--- program FrameL_C (robot ABB IRB 1300-10/1.15) ---
  Smooth(1)
  Set speed (1000.0 mm/s)
  Set Ref.: FrameL
  Set Tool: Generic Paint Sprayer
  Show Generic Paint Sprayer
  MoveJ 1 to (-1015.17, 960.31, 527.51) mm, rotated rx -115.53 ry -8.78 rz 162.28 deg; joints [74.023, 64.389, -177.634, 4.007, 86.75, 96.944, 1374.27, 3638.377, 370.799]
  MoveL 2 to (-1015.17, 960.31, 527.51) mm, rotated rx -115.53 ry -8.78 rz 162.28 deg; joints [74.023, 64.389, -177.634, 4.007, 86.75, 96.944, 1374.27, 3638.377, 370.799]
  MoveL 3 to (-1048.89, 876.36, 484.92) mm, rotated rx -115.53 ry -8.78 rz 162.28 deg; joints [74.023, 64.389, -177.634, 4.007, 86.75, 96.944, 1340.546, 3554.421, 413.392]
  MoveL 4 to (-1048.89, 876.36, 484.92) mm, rotated rx -115.53 ry -8.78 rz 162.28 deg; joints [74.023, 64.389, -177.634, 4.007, 86.75, 96.944, 1340.546, 3554.421, 413.392]
  Set speed (200.0 mm/s)
  MoveL 5 to (-1060.66, 876.62, 493.81) mm, rotated rx -115.95 ry -8.86 rz 162.43 deg; joints [74.023, 64.389, -177.634, 3.86, 86.355, 97.028, 1327.85, 3552.819, 401.035]
  MoveL 6 to (-1082.9, 876.62, 508.72) mm, rotated rx -117.21 ry -8.2 rz 164.5 deg; joints [74.023, 64.389, -177.634, 1.62, 85.639, 97.385, 1285.601, 3546.469, 378.721]
  MoveL 7 to (-1106.18, 876.62, 522.33) mm, rotated rx -120.93 ry -8.21 rz 166.59 deg; joints [74.023, 64.389, -177.634, -0.649, 82.446, 98.449, 1245.481, 3527.612, 337.393]
  MoveL 8 to (-1130.25, 876.36, 534.1) mm, rotated rx -123.9 ry -7.79 rz 168.6 deg; joints [74.023, 64.389, -177.635, -2.986, 80.093, 99.537, 1203.573, 3510.479, 305.654]
  MoveL 9 to (-1155.11, 876.1, 544.57) mm, rotated rx -126.6 ry -7.43 rz 170.12 deg; joints [74.023, 64.389, -179.794, -4.819, 80.083, 100.454, 1169.34, 3480.642, 285.56]
  MoveL 10 to (-1181.01, 875.83, 553.72) mm, rotated rx -129.64 ry -6.78 rz 171.9 deg; joints [74.023, 64.389, -182.144, -7.096, 80.08, 101.523, 1130.972, 3446.46, 267.382]
  MoveL 11 to (-1207.43, 875.31, 561.05) mm, rotated rx -132.01 ry -6.08 rz 173.29 deg; joints [74.023, 64.389, -183.913, -8.986, 80.08, 102.381, 1093.829, 3419.143, 254.394]
  MoveL 12 to (-1234.64, 874.79, 567.06) mm, rotated rx -134.1 ry -4.52 rz 175.35 deg; joints [74.023, 64.389, -185.084, -11.889, 80.08, 103.395, 1045.347, 3394.777, 245.717]
  MoveL 13 to (-1262.63, 874, 571.51) mm, rotated rx -135.78 ry -3.02 rz 177.06 deg; joints [74.023, 64.389, -185.959, -14.438, 80.08, 104.298, 998.548, 3373.942, 240.221]
  MoveL 14 to (-1290.62, 873.22, 574.39) mm, rotated rx -136.93 ry -1.36 rz 178.73 deg; joints [74.023, 64.389, -186.309, -16.976, 80.08, 105.132, 950.472, 3358.614, 238.296]
  MoveL 15 to (-1319.14, 872.43, 575.44) mm, rotated rx -138.23 ry 0.47 rz -179.58 deg; joints [74.023, 64.389, -186.628, -19.701, 79.974, 106.138, 900.949, 3341.306, 238.296]
  MoveL 16 to (-1347.65, 871.65, 574.39) mm, rotated rx -138.48 ry 3.29 rz -177.09 deg; joints [74.023, 64.389, -185.749, -23.502, 79.974, 107.295, 839.31, 3332.647, 245.735]
  MoveL 17 to (-1375.91, 870.6, 571.77) mm, rotated rx -138.43 ry 4.69 rz -175.85 deg; joints [74.023, 64.389, -185.157, -25.368, 79.974, 107.882, 794.724, 3328.918, 252.198]
  MoveL 18 to (-1403.9, 869.82, 567.06) mm, rotated rx -137.68 ry 7.29 rz -173.41 deg; joints [74.023, 64.389, -183.479, -28.797, 79.974, 108.923, 735.673, 3328.843, 265.904]
  MoveL 19 to (-1431.63, 868.77, 560.79) mm, rotated rx -136.77 ry 8.45 rz -172.14 deg; joints [74.023, 64.389, -182.957, -30.295, 80.608, 108.944, 693.869, 3328.843, 280.789]
  MoveL 20 to (-1458.84, 867.46, 552.68) mm, rotated rx -135.42 ry 10.6 rz -169.72 deg; joints [74.023, 64.389, -181.504, -33.244, 81.1, 109.501, 640.229, 3328.841, 301.523]
  MoveL 21 to (-1485.52, 866.15, 542.73) mm, rotated rx -133.88 ry 12.26 rz -167.55 deg; joints [74.023, 64.389, -180.635, -35.596, 82.031, 109.501, 592.858, 3327.208, 325.646]
  MoveL 22 to (-1511.42, 864.59, 530.96) mm, rotated rx -131.7 ry 14.03 rz -164.78 deg; joints [74.023, 64.389, -179.236, -38.372, 82.988, 109.462, 542.722, 3327.208, 354.62]
  MoveL 23 to (-1536.8, 862.75, 517.62) mm, rotated rx -129.53 ry 15.12 rz -162.45 deg; joints [74.023, 64.389, -178.191, -40.401, 83.978, 109.007, 499.686, 3327.208, 383.586]
  MoveL 24 to (-1560.87, 860.92, 502.71) mm, rotated rx -126.89 ry 16.3 rz -159.49 deg; joints [74.023, 64.389, -176.645, -42.942, 84.889, 108.635, 454.489, 3327.209, 416.346]
  MoveL 25 to (-1585.98, 858.31, 484.39) mm, rotated rx -125.12 ry 16.78 rz -157.68 deg; joints [74.023, 64.389, -175.535, -44.366, 85.349, 108.344, 417.425, 3327.209, 445.194]
  Set speed (1000.0 mm/s)
  MoveL 26 to (-1585.98, 858.31, 484.39) mm, rotated rx -125.12 ry 16.78 rz -157.68 deg; joints [74.023, 64.389, -175.535, -44.366, 85.349, 108.344, 417.425, 3327.209, 445.194]
  MoveL 27 to (-1632.41, 927.67, 539.47) mm, rotated rx -125.12 ry 16.78 rz -157.68 deg; joints [74.023, 64.389, -175.535, -44.366, 85.349, 108.344, 371.003, 3396.571, 390.114]
  Set speed (1000.0 mm/s)
  MoveL 28 to (-1782.13, 744.91, 885.74) mm, rotated rx -119.9 ry 6.95 rz -168.12 deg; joints [74.023, 82.832, -189.902, -29.809, 83.081, 103.224, 291.65, 3396.571, 197.643]
  MoveL 29 to (-1758.39, 661.31, 836.26) mm, rotated rx -119.9 ry 6.95 rz -168.12 deg; joints [74.023, 82.832, -189.902, -29.809, 83.081, 103.224, 315.396, 3312.976, 247.119]
  MoveL 30 to (-1758.39, 661.31, 836.26) mm, rotated rx -119.9 ry 6.95 rz -168.12 deg; joints [74.023, 82.832, -189.902, -29.809, 83.081, 103.224, 315.396, 3312.976, 247.119]
  Set speed (200.0 mm/s)
  MoveL 31 to (-1724.9, 670.47, 838.1) mm, rotated rx -121.18 ry 6.48 rz -169.44 deg; joints [74.023, 82.832, -191.204, -28.584, 83.081, 103.236, 361.581, 3315.861, 237.578]
  MoveL 32 to (-1691.68, 677.53, 839.67) mm, rotated rx -120.38 ry 5.33 rz -171 deg; joints [74.023, 82.942, -191.204, -26.541, 83.271, 102.399, 409.246, 3336.803, 237.579]
  MoveL 33 to (-1652.17, 686.16, 839.67) mm, rotated rx -120.13 ry 5.09 rz -171.3 deg; joints [74.023, 82.942, -191.058, -26.131, 83.271, 102.232, 451.408, 3349.272, 237.987]
  MoveL 34 to (-1610.05, 694.54, 839.67) mm, rotated rx -119.87 ry 4.65 rz -171.96 deg; joints [74.023, 82.942, -191.057, -25.301, 83.343, 101.933, 499.698, 3362.547, 237.986]
  MoveL 35 to (-1562.18, 702.65, 839.67) mm, rotated rx -119.38 ry 4.09 rz -172.77 deg; joints [74.023, 82.942, -190.802, -24.26, 83.343, 101.565, 554.808, 3378.986, 238.548]
  MoveL 36 to (-1528.43, 707.88, 839.4) mm, rotated rx -119.36 ry 3.58 rz -173.66 deg; joints [74.023, 82.942, -190.956, -23.231, 83.343, 101.335, 597.012, 3388.041, 237.249]
  MoveL 37 to (-1485.26, 713.63, 838.88) mm, rotated rx -118.87 ry 2.94 rz -174.68 deg; joints [74.023, 82.942, -190.736, -21.967, 83.343, 100.942, 649.473, 3402.601, 238.129]
  MoveL 38 to (-1441.83, 719.13, 838.1) mm, rotated rx -117.68 ry 2.67 rz -174.93 deg; joints [74.023, 82.942, -189.774, -21.484, 83.343, 100.534, 693.898, 3420.583, 243.983]
  MoveL 39 to (-1401.81, 723.58, 837.57) mm, rotated rx -117.2 ry 2.44 rz -175.26 deg; joints [74.023, 82.942, -189.426, -21.034, 83.343, 100.319, 736.495, 3430.885, 246.249]
  MoveL 40 to (-1370.15, 726.98, 837.05) mm, rotated rx -116.96 ry 2.24 rz -175.61 deg; joints [74.023, 82.942, -189.285, -20.596, 83.343, 100.172, 771.246, 3437.889, 247.356]
  MoveL 41 to (-1348.7, 729.07, 836.53) mm, rotated rx -116.25 ry 1.82 rz -176.31 deg; joints [74.023, 82.942, -188.793, -19.705, 83.343, 99.816, 798.461, 3449.363, 250.333]
  MoveL 42 to (-1313.64, 732.47, 835.74) mm, rotated rx -115.78 ry 1.8 rz -176.28 deg; joints [74.023, 82.942, -188.382, -19.671, 83.343, 99.686, 832.592, 3457.166, 253.563]
  MoveL 43 to (-1272.05, 736.66, 834.7) mm, rotated rx -115.78 ry 1.8 rz -176.28 deg; joints [74.023, 82.942, -188.382, -19.671, 83.343, 99.686, 874.188, 3461.352, 254.61]
  Set speed (1000.0 mm/s)
  MoveL 44 to (-1272.05, 736.66, 834.7) mm, rotated rx -115.78 ry 1.8 rz -176.28 deg; joints [74.023, 82.942, -188.382, -19.671, 83.343, 99.686, 874.188, 3461.352, 254.61]
  MoveL 45 to (-1279.25, 826.43, 878.16) mm, rotated rx -115.78 ry 1.8 rz -176.28 deg; joints [74.023, 82.942, -188.382, -19.671, 83.343, 99.686, 866.984, 3551.122, 211.142]
  Set speed (1000.0 mm/s)
  MoveL 46 to (-1224.09, 625.8, 1224.25) mm, rotated rx -153.49 ry 17.59 rz -171.43 deg; joints [74.023, 113.295, -210, -50.489, 58.121, 141.888, 800.056, 3107.358, 0]
  MoveL 47 to (-1190.69, 585.7, 1138.95) mm, rotated rx -153.49 ry 17.59 rz -171.43 deg; joints [74.023, 113.295, -210, -50.489, 58.121, 141.888, 833.458, 3067.258, 85.301]
  MoveL 48 to (-1190.69, 585.7, 1138.95) mm, rotated rx -153.49 ry 17.59 rz -171.43 deg; joints [74.023, 113.295, -210, -50.489, 58.121, 141.888, 833.458, 3067.258, 85.301]
  Set speed (200.0 mm/s)
  MoveL 49 to (-1213.18, 590.41, 1127.7) mm, rotated rx -152.92 ry 17.68 rz -171.17 deg; joints [74.109, 113.295, -209.797, -50.489, 58.34, 141.571, 810.153, 3076.307, 98.867]
  MoveL 50 to (-1232.02, 595.91, 1115.67) mm, rotated rx -149.63 ry 20.03 rz -168.65 deg; joints [74.109, 113.295, -209.797, -51.349, 61.878, 139.926, 770.209, 3087.414, 138.308]
  MoveL 51 to (-1245.36, 601.66, 1104.16) mm, rotated rx -144.68 ry 22.57 rz -164.79 deg; joints [74.109, 113.295, -209.797, -52.484, 66.425, 137.222, 731.825, 3098.93, 187.325]
  MoveL 52 to (-1255.57, 608.2, 1091.34) mm, rotated rx -138.48 ry 23.76 rz -160.37 deg; joints [74.109, 113.295, -209.797, -53.093, 70.737, 133.096, 702.117, 3113.993, 238.067]
  MoveL 53 to (-1266.03, 615.79, 1076.43) mm, rotated rx -135.62 ry 23.47 rz -158.71 deg; joints [74.355, 113.295, -209.797, -53.093, 72.19, 130.762, 689.721, 3129.009, 266.528]
  MoveL 54 to (-1277.02, 624.69, 1059.16) mm, rotated rx -132.74 ry 23.27 rz -156.85 deg; joints [74.355, 113.295, -209.797, -53.171, 73.8, 128.56, 673.065, 3142.176, 298.917]
  MoveL 55 to (-1289.58, 634.63, 1039.02) mm, rotated rx -131.52 ry 23.24 rz -155.98 deg; joints [74.355, 113.295, -209.797, -53.335, 74.526, 127.689, 657.589, 3152.866, 325.984]
  MoveL 56 to (-1302.66, 645.09, 1016.52) mm, rotated rx -130.52 ry 22.58 rz -155.81 deg; joints [74.946, 113.295, -209.797, -53.335, 74.692, 126.502, 651.96, 3170.749, 350.648]
  MoveL 57 to (-1314.95, 656.34, 992.97) mm, rotated rx -127.95 ry 21.97 rz -154.38 deg; joints [75.07, 113.295, -209.797, -53.335, 75.943, 124.315, 637.676, 3187.198, 386.491]
  MoveL 58 to (-1325.16, 667.33, 969.69) mm, rotated rx -124.78 ry 21.2 rz -152.49 deg; joints [75.07, 113.295, -209.797, -53.423, 77.573, 121.661, 622.718, 3202.179, 425.966]
  MoveL 59 to (-1331.7, 677.01, 948.5) mm, rotated rx -121.28 ry 19.57 rz -151.13 deg; joints [75.729, 113.295, -209.797, -53.423, 78.977, 118.19, 621.847, 3223.413, 462.069]
  MoveL 60 to (-1334.83, 686.16, 929.14) mm, rotated rx -115.7 ry 16.94 rz -148.81 deg; joints [76.214, 113.295, -209.797, -53.423, 81.501, 112.732, 620.29, 3244.805, 508.191]
  MoveL 61 to (-1335.36, 694.54, 911.09) mm, rotated rx -112.21 ry 15.04 rz -147.57 deg; joints [76.419, 113.295, -209.796, -53.344, 83.103, 109.182, 620.29, 3260.09, 543.538]
  MoveL 62 to (-1334.05, 702.65, 894.34) mm, rotated rx -108.35 ry 12.58 rz -146.71 deg; joints [76.419, 113.295, -208.835, -52.795, 84.285, 105.811, 620.291, 3284.293, 577.893]
  MoveL 63 to (-1330.91, 710.23, 878.65) mm, rotated rx -106.25 ry 11.06 rz -146.65 deg; joints [76.419, 113.295, -207.305, -52.247, 84.285, 104.649, 622.688, 3310.154, 601.765]
  MoveL 64 to (-1326.72, 717.82, 863.73) mm, rotated rx -104 ry 9.39 rz -146.81 deg; joints [76.419, 113.295, -205.674, -51.514, 84.285, 103.354, 626.889, 3338.129, 626.047]
  MoveL 65 to (-1321.23, 725.14, 849.35) mm, rotated rx -102.7 ry 8.13 rz -147.88 deg; joints [76.419, 113.295, -204.934, -50.104, 84.286, 102.209, 637.653, 3363.4, 645.188]
  MoveL 66 to (-1354.46, 721.74, 850.39) mm, rotated rx -175.54 ry 33.28 rz 101.98 deg; joints [56.988, 143.589, -137.16, 144.417, 41.145, 36.117, 651.946, 3698.807, 1100]
  MoveL 67 to (-1365.71, 720.44, 850.65) mm, rotated rx -146.28 ry 2.17 rz -178.55 deg; joints [76.42, 113.126, -204.934, -34.5, 46.983, 127.515, 802.993, 3345.808, 316.76]
  MoveL 68 to (-1402.07, 716.25, 851.7) mm, rotated rx -146.28 ry 2.15 rz -178.57 deg; joints [76.452, 113.127, -204.934, -34.5, 46.968, 127.491, 767.195, 3341.791, 315.632]
  MoveL 69 to (-1441.57, 711.54, 852.75) mm, rotated rx -147.29 ry 2.97 rz -178.09 deg; joints [76.452, 113.127, -205.051, -36.188, 46.968, 129.159, 719.979, 3326.698, 313.434]
  MoveL 70 to (-1483.95, 705.52, 854.05) mm, rotated rx -147.72 ry 2.66 rz -178.32 deg; joints [76.657, 113.126, -205.225, -36.188, 46.589, 129.171, 683.277, 3317.897, 308.963]
  MoveL 71 to (-1526.07, 699.25, 855.1) mm, rotated rx -148.75 ry 3.4 rz -177.94 deg; joints [76.657, 113.126, -205.394, -37.74, 46.589, 130.742, 634.518, 3301.013, 306.662]
  MoveL 72 to (-1565.32, 692.97, 855.89) mm, rotated rx -149.59 ry 4.5 rz -177.37 deg; joints [76.657, 113.076, -205.394, -39.637, 46.907, 132.518, 585.134, 3285.408, 306.662]
  MoveL 73 to (-1604.04, 685.64, 856.67) mm, rotated rx -149.63 ry 4.75 rz -177.22 deg; joints [76.657, 113.053, -205.394, -39.955, 47.091, 132.754, 544.052, 3276.943, 306.662]
  MoveL 74 to (-1644.85, 677.27, 857.19) mm, rotated rx -149.67 ry 5.03 rz -177.07 deg; joints [76.657, 112.983, -205.394, -40.272, 47.328, 132.968, 500.693, 3267.189, 306.662]
  MoveL 75 to (-1683.3, 668.64, 857.72) mm, rotated rx -149.88 ry 4.86 rz -177.19 deg; joints [76.768, 112.983, -205.475, -40.272, 47.126, 132.968, 465.246, 3257.352, 304.541]
  MoveL 76 to (-1714.44, 661.05, 857.72) mm, rotated rx -150.07 ry 5.32 rz -176.94 deg; joints [76.768, 112.823, -205.475, -40.855, 47.48, 133.411, 429.986, 3246.468, 304.541]
  MoveL 77 to (-1699.79, 652.15, 878.91) mm, rotated rx -108.33 ry -41.93 rz 178.16 deg; joints [107.262, 119.949, -159.707, -81.239, 23.985, 121.042, 1096.293, 3778.444, 604.845]
  MoveL 78 to (-1684.35, 642.74, 900.88) mm, rotated rx -103.77 ry -3.13 rz 167.42 deg; joints [76.148, 112.823, -205.475, -3.654, 79.163, 94.041, 621.106, 3510.146, 535.977]
  MoveL 79 to (-1667.87, 633.06, 924.17) mm, rotated rx -103.52 ry -3.2 rz 166.93 deg; joints [76.148, 113.008, -205.475, -3.137, 79.163, 93.889, 642.032, 3502.509, 516.04]
  MoveL 80 to (-1650.34, 622.85, 949.02) mm, rotated rx -103.61 ry -3.24 rz 166.87 deg; joints [76.148, 113.007, -205.475, -3.08, 79.072, 93.904, 660.131, 3492.212, 490.338]
  MoveL 81 to (-1668.13, 617.1, 950.85) mm, rotated rx -150.18 ry 3.36 rz -178.08 deg; joints [76.148, 127.331, -159.488, -126.409, 33.343, 234.838, 410.502, 3521.9, 490.338]
  MoveL 82 to (-1646.94, 607.16, 976.49) mm, rotated rx -103.2 ry -21.92 rz 173.54 deg; joints [79.337, 132.004, -146.722, -134.913, 10.128, 208.962, 623.21, 3814.134, 838.601]
  MoveL 83 to (-1626.27, 597.74, 1000.82) mm, rotated rx -103.03 ry 17 rz 164.34 deg; joints [83.994, 114.805, -210, -10.723, 92.781, 110.214, 765.634, 3467.741, 546.847]
  MoveL 84 to (-1604.3, 587.54, 1026.46) mm, rotated rx -102.27 ry -2.64 rz 168.02 deg; joints [68.793, 127.331, -142.872, 39.964, 4.671, 54.643, 479.375, 3792.466, 820.793]
  MoveL 85 to (-1591.22, 581.26, 1041.37) mm, rotated rx -102.7 ry -2.7 rz 168.18 deg; joints [68.793, 127.33, -143.048, 40.106, 4.387, 54.643, 491.326, 3784.586, 800.784]
  MoveL 86 to (-1576.3, 574.19, 1058.38) mm, rotated rx -102.74 ry -2.72 rz 168.15 deg; joints [68.821, 127.318, -143.074, 40.113, 4.387, 54.643, 506.991, 3777.652, 783.064]
  MoveL 87 to (-1558.25, 565.82, 1078.78) mm, rotated rx -102.36 ry -3.02 rz 166.5 deg; joints [69.84, 127.318, -143.735, 40.113, 5.465, 54.375, 557.879, 3777.653, 760.069]
  MoveL 88 to (-1552.24, 562.68, 1085.58) mm, rotated rx -103.74 ry -3.73 rz 165.11 deg; joints [71.265, 127.318, -145.275, 40.29, 5.465, 54.375, 602.999, 3777.836, 728.411]
  MoveL 89 to (-1529.74, 549.6, 1110.17) mm, rotated rx -104.95 ry -3.95 rz 165.55 deg; joints [71.265, 127.318, -145.818, 40.635, 4.699, 54.375, 622.506, 3759.732, 689.247]
  MoveL 90 to (-1522.15, 545.15, 1118.55) mm, rotated rx -106.77 ry -4.5 rz 165.41 deg; joints [71.357, 127.318, -147.645, 41.199, 4.699, 54.375, 636.151, 3745.82, 651.363]
  MoveL 91 to (-1514.83, 540.71, 1126.66) mm, rotated rx -108.15 ry -4.97 rz 165.21 deg; joints [71.531, 127.318, -149.051, 41.589, 4.699, 54.375, 650.887, 3734.192, 620.842]
  MoveL 92 to (-1509.07, 536.52, 1132.93) mm, rotated rx -109.08 ry -4.93 rz 166.05 deg; joints [71.623, 127.66, -149.051, 41.589, 3.22, 54.557, 650.887, 3725.698, 612.176]
  MoveL 93 to (-1479.25, 539.4, 1137.12) mm, rotated rx -96.71 ry 0.66 rz -174.4 deg; joints [52.115, 127.659, -135.62, 39.626, 3.22, 54.557, 184.512, 3559.834, 826.74]
  MoveL 94 to (-1446.02, 542.02, 1141.57) mm, rotated rx -96.9 ry 0.66 rz -174.6 deg; joints [52.293, 127.659, -135.786, 39.725, 3.22, 54.557, 222.003, 3564.9, 819.431]
  MoveL 95 to (-1405.47, 545.15, 1147.32) mm, rotated rx -96.24 ry 0.57 rz -174.82 deg; joints [52.145, 127.685, -135.786, 39.725, 3.877, 54.18, 262.446, 3568.064, 819.43]
  MoveL 96 to (-1359.69, 548.56, 1153.34) mm, rotated rx -95.72 ry 0.46 rz -175.39 deg; joints [52.145, 127.685, -136.116, 39.725, 4.814, 53.897, 313.297, 3574.124, 815.026]
  MoveL 97 to (-1311.03, 551.96, 1159.88) mm, rotated rx -93.84 ry 0.28 rz -175.81 deg; joints [51.521, 127.643, -136.116, 38.704, 6.754, 53.892, 356.743, 3574.124, 823.22]
  MoveL 98 to (-1261.84, 555.1, 1165.9) mm, rotated rx -94.32 ry 0.29 rz -176.15 deg; joints [51.809, 127.643, -136.507, 38.986, 6.754, 53.892, 413.141, 3581.111, 810.29]
  MoveL 99 to (-1215.02, 557.97, 1171.39) mm, rotated rx -92.6 ry 0.13 rz -177.14 deg; joints [51.285, 127.075, -136.507, 38.986, 9.273, 53.02, 459.516, 3585.376, 810.29]
  MoveL 100 to (-1166.36, 560.59, 1176.62) mm, rotated rx -90.9 ry 0.05 rz -177.14 deg; joints [50.926, 127.075, -135.847, 37.989, 10.12, 53.02, 502.442, 3585.376, 824.087]
  MoveL 101 to (-1111.42, 562.94, 1181.86) mm, rotated rx -88.74 ry -0.04 rz -178.11 deg; joints [50.117, 126.225, -135.847, 37.074, 13.323, 52.861, 552.192, 3585.376, 824.096]
  MoveL 102 to (-1049.68, 565.56, 1187.09) mm, rotated rx -86.59 ry -0.11 rz -178.18 deg; joints [49.822, 126.225, -134.979, 35.766, 14.298, 52.861, 609.4, 3585.372, 843.363]
  MoveL 103 to (-981.39, 567.91, 1192.32) mm, rotated rx -85.14 ry -0.19 rz -177.72 deg; joints [49.495, 126.224, -133.896, 34.792, 14.298, 52.861, 668.023, 3582.496, 858.047]
  MoveL 104 to (-904.48, 570.79, 1197.55) mm, rotated rx -82.67 ry -0.17 rz -178.69 deg; joints [48.935, 125.631, -133.896, 33.479, 17.36, 52.86, 743.872, 3582.496, 864.961]
  MoveL 105 to (-818.15, 573.41, 1202.52) mm, rotated rx -79.46 ry -0.27 rz -178.56 deg; joints [48.899, 125.631, -131.755, 31.359, 17.672, 52.86, 826.261, 3582.495, 902.412]
  MoveL 106 to (-727.89, 576.29, 1206.71) mm, rotated rx -76.16 ry -0.16 rz -179.35 deg; joints [48.815, 125.631, -130.971, 29.412, 19.77, 52.86, 921.427, 3582.494, 932.118]
  MoveL 107 to (-639.73, 578.9, 1209.85) mm, rotated rx -75.2 ry -0.12 rz -179.54 deg; joints [48.665, 125.631, -130.915, 28.851, 20.562, 52.86, 1009.092, 3582.084, 937.49]
  MoveL 108 to (-560.72, 581.26, 1212.2) mm, rotated rx -74.25 ry -0.19 rz -179.34 deg; joints [48.251, 125.631, -130.748, 28.203, 21.141, 52.86, 1080.603, 3576.71, 943.985]
  MoveL 109 to (-498.72, 583.09, 1213.25) mm, rotated rx -72.59 ry -0.34 rz -178.92 deg; joints [47.368, 125.631, -130.664, 27.035, 22.339, 52.86, 1126.833, 3562.073, 956.627]
  MoveL 110 to (-447.18, 584.66, 1213.25) mm, rotated rx -73.06 ry -0.49 rz -178.38 deg; joints [47.122, 125.631, -130.664, 27.035, 21.798, 53.038, 1170.327, 3559.537, 952.194]
  MoveL 111 to (-400.61, 585.97, 1212.73) mm, rotated rx -72.12 ry -0.65 rz -177.98 deg; joints [46.48, 125.631, -130.66, 26.321, 22.465, 53.038, 1204.822, 3548.789, 959.813]
  MoveL 112 to (-356.92, 587.54, 1211.94) mm, rotated rx -70.24 ry -0.72 rz -177.99 deg; joints [45.923, 125.631, -130.659, 25.065, 23.969, 53.038, 1241.071, 3538.165, 975.631]
  MoveL 113 to (-315.06, 588.84, 1210.63) mm, rotated rx -70.43 ry -0.9 rz -177.46 deg; joints [45.525, 125.631, -130.659, 25.049, 23.68, 53.038, 1273.107, 3532.715, 974.676]
  MoveL 114 to (-272.42, 590.41, 1208.8) mm, rotated rx -70.97 ry -0.97 rz -177.19 deg; joints [45.384, 125.631, -130.79, 25.348, 23.331, 53.038, 1311.73, 3532.716, 970.896]
  MoveL 115 to (-226.9, 591.98, 1206.45) mm, rotated rx -73.64 ry -0.96 rz -176.74 deg; joints [44.998, 125.631, -132.354, 27.122, 22.863, 53.038, 1350.313, 3532.716, 940.01]
  MoveL 116 to (-177.19, 594.08, 1203.57) mm, rotated rx -73.35 ry -0.99 rz -176.7 deg; joints [44.899, 125.631, -132.32, 26.914, 23.048, 53.038, 1398.384, 3532.716, 945.435]
  MoveL 117 to (-122.25, 596.95, 1199.65) mm, rotated rx -71 ry -1.16 rz -176.62 deg; joints [44.814, 125.631, -130.978, 25.227, 23.367, 53.038, 1449.764, 3529.34, 977.622]
  MoveL 118 to (-64.7, 600.35, 1194.68) mm, rotated rx -71.58 ry -1.55 rz -175.36 deg; joints [43.91, 125.631, -130.978, 25.227, 22.594, 53.107, 1484.953, 3516.791, 976.338]
  MoveL 119 to (-7.41, 604.28, 1188.4) mm, rotated rx -71.84 ry -2 rz -173.91 deg; joints [42.65, 125.483, -130.978, 25.042, 22.207, 53.107, 1513.724, 3498.226, 976.338]
  MoveL 120 to (47.53, 608.73, 1180.55) mm, rotated rx -71.95 ry -2.25 rz -173.12 deg; joints [41.878, 125.238, -130.978, 24.927, 22.207, 53.107, 1551.811, 3489.375, 978.496]
  MoveL 121 to (97.76, 613.17, 1171.39) mm, rotated rx -72.14 ry -2.58 rz -172.05 deg; joints [40.827, 124.881, -130.978, 24.806, 22.207, 53.107, 1579.348, 3475.469, 979.235]
  MoveL 122 to (146.16, 618.14, 1160.67) mm, rotated rx -71.66 ry -3.12 rz -170.66 deg; joints [39.492, 124.881, -130.973, 24.071, 22.208, 53.107, 1600.414, 3453.1, 991.733]
  MoveL 123 to (195.08, 623.9, 1148.11) mm, rotated rx -70.72 ry -3.9 rz -168.99 deg; joints [37.886, 124.881, -130.779, 22.861, 22.208, 53.107, 1616.753, 3424.083, 1010.129]
  MoveL 124 to (244.27, 630.96, 1132.67) mm, rotated rx -72.37 ry -4.39 rz -166.45 deg; joints [36.316, 124.881, -130.779, 22.861, 20.403, 53.762, 1629.557, 3398.061, 1010.086]
  MoveL 125 to (293.45, 639.6, 1113.05) mm, rotated rx -73.81 ry -4.79 rz -163.94 deg; joints [34.487, 124.485, -130.779, 22.861, 19.275, 54.345, 1640.022, 3368.784, 1010.086]
  MoveL 126 to (347.34, 650.58, 1088.98) mm, rotated rx -75.56 ry -4.41 rz -163.38 deg; joints [33.9, 124.103, -131.5, 24.28, 19.275, 54.345, 1684.493, 3372.016, 1010.086]
  MoveL 127 to (411.18, 663.4, 1059.94) mm, rotated rx -77.83 ry -3.62 rz -163.67 deg; joints [34.059, 123.592, -132.235, 26.347, 19.275, 54.345, 1752.616, 3394.507, 1010.086]
  MoveL 128 to (478.41, 677.27, 1028.03) mm, rotated rx -76.13 ry -4.13 rz -163.75 deg; joints [33.354, 123.589, -132.235, 25.979, 20.539, 53.289, 1812.432, 3394.507, 1054.104]
  MoveL 129 to (541.98, 690.61, 996.11) mm, rotated rx -77.3 ry -3.78 rz -163.69 deg; joints [32.777, 122.082, -132.235, 27.086, 21.487, 53.29, 1865.951, 3404.149, 1054.105]
  MoveL 130 to (598.49, 702.38, 966.55) mm, rotated rx -81.33 ry -2.4 rz -164.67 deg; joints [33.246, 122.082, -134.352, 30.848, 21.487, 53.29, 1939.65, 3433.922, 1040.16]
  MoveL 131 to (643.49, 711.8, 942.22) mm, rotated rx -81.55 ry -2.4 rz -164.23 deg; joints [32.765, 121.878, -134.352, 30.997, 21.523, 53.29, 1976.214, 3433.922, 1059.38]
  MoveL 132 to (682.21, 719.91, 920.5) mm, rotated rx -82.28 ry -2.2 rz -164.16 deg; joints [32.181, 120.834, -134.352, 31.735, 22.267, 53.29, 2006.381, 3435.187, 1059.38]
  MoveL 133 to (719.36, 727.76, 899.05) mm, rotated rx -81.72 ry -2.4 rz -163.96 deg; joints [31.793, 120.699, -134.352, 31.309, 22.767, 53.248, 2037.804, 3435.187, 1082.681]
  MoveL 134 to (754.41, 735.09, 878.65) mm, rotated rx -79.11 ry -3.34 rz -163.15 deg; joints [31.295, 117.378, -129.937, 28.826, 23.013, 53.248, 2045.276, 3435.187, 1100]
  MoveL 135 to (786.59, 741.63, 859.03) mm, rotated rx -81.68 ry -2.48 rz -163.48 deg; joints [31.207, 117.378, -131.27, 31.246, 23.013, 53.248, 2082.657, 3444.94, 1091.877]
  MoveL 136 to (817.2, 748.17, 839.93) mm, rotated rx -80.71 ry -2.91 rz -162.77 deg; joints [30.689, 115.081, -128.534, 30.247, 23.013, 53.248, 2093.261, 3443.042, 1100]
  MoveL 137 to (846.24, 754.18, 821.61) mm, rotated rx -82.59 ry -2.12 rz -164.12 deg; joints [31.66, 115.081, -129.394, 32.148, 23.013, 53.248, 2143.77, 3474.649, 1099.433]
  MoveL 138 to (874.76, 760.2, 803.3) mm, rotated rx -81.97 ry -2.36 rz -163.7 deg; joints [31.181, 112.683, -126.999, 31.58, 23.359, 53.248, 2156.086, 3474.648, 1100]
  Set speed (1000.0 mm/s)
  MoveL 139 to (874.76, 760.2, 803.3) mm, rotated rx -81.97 ry -2.36 rz -163.7 deg; joints [31.181, 112.683, -126.999, 31.58, 23.359, 53.248, 2156.086, 3474.648, 1100]
  MoveL 140 to (846.41, 855.08, 789.34) mm, rotated rx -81.97 ry -2.36 rz -163.7 deg; joints [30.702, 111.825, -126.999, 31.58, 24.332, 53.381, 2122.171, 3562.297, 1100]
  Set speed (1000.0 mm/s)
  MoveL 141 to (1541.36, 940.82, 613.61) mm, rotated rx -125.26 ry -7.23 rz 169.91 deg; joints [30.702, 111.825, -161.462, 74.993, 31.83, 53.381, 3191.702, 3594.263, 705.738]
  MoveL 142 to (1519.9, 861.71, 556.34) mm, rotated rx -125.26 ry -7.23 rz 169.91 deg; joints [30.702, 111.825, -161.462, 74.992, 31.83, 53.381, 3170.245, 3515.153, 763.012]
  MoveL 143 to (1519.9, 861.71, 556.34) mm, rotated rx -125.26 ry -7.23 rz 169.91 deg; joints [30.702, 111.825, -161.462, 74.992, 31.83, 53.381, 3170.245, 3515.153, 763.012]
  Set speed (200.0 mm/s)
  MoveL 144 to (1494, 861.45, 566.8) mm, rotated rx -125.78 ry -6.92 rz 170.51 deg; joints [30.702, 112.149, -161.462, 74.964, 31.003, 53.381, 3137.514, 3511.708, 754.412]
  MoveL 145 to (1489.29, 872.43, 551.89) mm, rotated rx -123.78 ry -6.41 rz 170.52 deg; joints [29.063, 112.149, -160.887, 74.915, 33.272, 53.381, 3113.809, 3511.71, 787.542]
  MoveL 146 to (1461.56, 872.96, 561.57) mm, rotated rx -124.95 ry -6.3 rz 171.08 deg; joints [29.508, 112.243, -160.887, 75.006, 31.785, 53.381, 3084.564, 3511.71, 771.24]
  MoveL 147 to (1433.04, 873.48, 569.68) mm, rotated rx -126.07 ry -5.47 rz 172.55 deg; joints [29.508, 113.123, -160.887, 74.89, 29.817, 53.381, 3039.121, 3504.629, 770.22]
  MoveL 148 to (1404.52, 874.26, 576.22) mm, rotated rx -127.67 ry -4.4 rz 174.32 deg; joints [29.608, 114.1, -160.812, 74.89, 27.168, 53.381, 2990.793, 3495.601, 770.22]
  MoveL 149 to (1375.22, 875.05, 580.67) mm, rotated rx -128.32 ry -3.5 rz 175.58 deg; joints [29.609, 114.229, -159.976, 74.684, 25.574, 53.381, 2943.185, 3492.131, 770.22]
  MoveL 150 to (1345.92, 876.1, 583.81) mm, rotated rx -128.52 ry -2.35 rz 177.05 deg; joints [29.609, 114.229, -158.608, 74.132, 24.01, 53.381, 2890.52, 3491.681, 776.48]
  MoveL 151 to (1316.1, 876.88, 585.12) mm, rotated rx -127.31 ry -1.42 rz 178.14 deg; joints [29.1, 114.229, -157.227, 73.229, 24.008, 53.381, 2837.13, 3491.681, 793.636]
  MoveL 152 to (1286.01, 877.67, 585.38) mm, rotated rx -125.42 ry -0.49 rz 179.31 deg; joints [28.402, 114.229, -155.682, 71.968, 24.501, 53.381, 2781.001, 3491.681, 817.801]
  MoveL 153 to (1255.14, 878.45, 584.07) mm, rotated rx -122.83 ry 0.38 rz -179.41 deg; joints [27.568, 114.229, -154.001, 70.247, 25.437, 53.381, 2722.233, 3491.682, 849.706]
  MoveL 154 to (1223.49, 879.24, 581.45) mm, rotated rx -120.01 ry 0.77 rz -178.66 deg; joints [26.72, 114.229, -152.909, 68.545, 27.094, 53.381, 2671.668, 3491.684, 880.366]
  MoveL 155 to (1190.26, 879.5, 578.05) mm, rotated rx -117.18 ry 1.29 rz -177.49 deg; joints [26.075, 114.229, -151.527, 66.485, 28.178, 53.381, 2616.373, 3491.684, 914.661]
  MoveL 156 to (1155.47, 879.5, 573.87) mm, rotated rx -116.01 ry 1.07 rz -177.82 deg; joints [26.075, 114.16, -151.527, 65.79, 29.242, 53.381, 2584.953, 3497.655, 925.992]
  MoveL 157 to (1117.01, 879.24, 569.16) mm, rotated rx -111.18 ry 0.83 rz -177.85 deg; joints [24.971, 114.161, -151.225, 63.037, 33.256, 53.381, 2537.979, 3497.655, 969.43]
  MoveL 158 to (1107.07, 868.25, 594.8) mm, rotated rx -116 ry 0.51 rz -178.95 deg; joints [26.602, 114.161, -152.303, 65.955, 29.946, 53.381, 2554.828, 3497.655, 898.648]
  MoveL 159 to (1106.28, 861.97, 607.09) mm, rotated rx -118.35 ry 0.15 rz -179.73 deg; joints [27.54, 114.16, -153.145, 67.339, 28.498, 53.381, 2572.558, 3497.655, 862.408]
  MoveL 160 to (1067.3, 855.17, 619.65) mm, rotated rx -120.95 ry -0.25 rz 179.58 deg; joints [28.69, 114.16, -154.04, 68.676, 26.683, 53.381, 2553.898, 3497.655, 824.139]
  MoveL 161 to (1017.6, 845.23, 638.48) mm, rotated rx -122.6 ry -1.12 rz 178.25 deg; joints [29.774, 114.16, -155.4, 69.641, 26.174, 53.381, 2533.298, 3497.655, 782.834]
  MoveL 162 to (977.57, 845.23, 640.58) mm, rotated rx -121.89 ry -1.11 rz 178.22 deg; joints [29.525, 114.16, -155.285, 69.349, 26.819, 53.381, 2490.792, 3497.658, 786.521]
  MoveL 163 to (935.97, 845.23, 643.19) mm, rotated rx -121.07 ry -1.09 rz 178.19 deg; joints [29.243, 114.16, -155.155, 69, 27.567, 53.381, 2446.403, 3497.658, 790.674]
  MoveL 164 to (924.99, 833.19, 664.12) mm, rotated rx -120.71 ry -1.09 rz 178.17 deg; joints [29.523, 114.331, -155.154, 68.587, 27.563, 53.381, 2437.619, 3491.47, 774.824]
  MoveL 165 to (917.4, 825.08, 678.25) mm, rotated rx -120.01 ry -1.07 rz 178.15 deg; joints [29.835, 114.949, -155.154, 68.534, 27.625, 52.692, 2432.154, 3491.47, 774.824]
  MoveL 166 to (912.43, 820.11, 687.93) mm, rotated rx -118.12 ry -1.03 rz 178.08 deg; joints [29.552, 114.949, -154.763, 67.478, 29.028, 52.692, 2423.355, 3491.494, 781.508]
  MoveL 167 to (907.98, 815.92, 696.56) mm, rotated rx -117.18 ry -1 rz 178.05 deg; joints [29.536, 114.97, -154.56, 66.865, 29.626, 52.692, 2417.985, 3491.495, 781.508]
  MoveL 168 to (945.13, 815.66, 693.69) mm, rotated rx -117.42 ry -1.01 rz 178.05 deg; joints [29.536, 114.896, -154.56, 66.994, 29.486, 52.723, 2455.16, 3490.236, 781.508]
  MoveL 169 to (982.02, 815.4, 690.81) mm, rotated rx -117.89 ry -1.02 rz 178.07 deg; joints [29.696, 114.896, -154.623, 67.203, 29.06, 52.723, 2493.6, 3490.236, 780.424]
  MoveL 170 to (1018.91, 815.14, 688.19) mm, rotated rx -118.36 ry -1.23 rz 177.73 deg; joints [29.832, 114.896, -155.009, 67.591, 29.016, 52.723, 2536.911, 3490.235, 776.618]
  MoveL 171 to (1056.05, 814.62, 685.31) mm, rotated rx -119.54 ry -1.67 rz 177.06 deg; joints [30.199, 114.896, -155.82, 68.447, 28.69, 52.723, 2587.894, 3490.23, 764.715]
  MoveL 172 to (1094.51, 814.09, 682.17) mm, rotated rx -120.25 ry -1.69 rz 177.1 deg; joints [30.472, 114.896, -155.921, 68.72, 28.018, 52.723, 2628.94, 3490.229, 761.976]
  MoveL 173 to (1134.8, 813.31, 678.77) mm, rotated rx -120.96 ry -1.71 rz 177.15 deg; joints [30.769, 114.896, -156.022, 68.974, 27.328, 52.723, 2672.03, 3490.229, 759.546]
  MoveL 174 to (1177.97, 812.52, 674.85) mm, rotated rx -121.67 ry -2.16 rz 176.51 deg; joints [31.045, 114.896, -156.75, 69.55, 27.334, 52.723, 2727.821, 3490.229, 752.808]
  MoveL 175 to (1222.44, 811.48, 670.66) mm, rotated rx -121.68 ry -2.37 rz 176.17 deg; joints [31.073, 114.693, -156.846, 69.689, 27.649, 52.723, 2776.774, 3490.229, 752.808]
  MoveL 176 to (1266.65, 810.43, 666.22) mm, rotated rx -121.92 ry -2.59 rz 175.86 deg; joints [31.218, 114.666, -157.142, 69.894, 27.703, 52.723, 2827.021, 3490.229, 752.808]
  MoveL 177 to (1308.77, 809.12, 661.51) mm, rotated rx -124.52 ry -2.92 rz 175.77 deg; joints [32.313, 114.666, -157.886, 70.872, 25.463, 52.723, 2884.542, 3490.151, 733.89]
  MoveL 178 to (1347.49, 807.81, 657.32) mm, rotated rx -125.02 ry -3.6 rz 174.87 deg; joints [32.613, 114.666, -158.852, 71.389, 25.852, 52.723, 2940.606, 3490.151, 727.32]
  MoveL 179 to (1385.95, 806.24, 652.35) mm, rotated rx -125.03 ry -3.83 rz 174.56 deg; joints [32.686, 114.384, -158.852, 71.49, 26.104, 52.723, 2983.535, 3490.151, 727.478]
  MoveL 180 to (1427.28, 804.15, 646.59) mm, rotated rx -125.23 ry -4.17 rz 174.12 deg; joints [32.909, 114.274, -159.19, 71.666, 26.266, 52.723, 3033.678, 3490.151, 727.478]
  MoveL 181 to (1486.67, 800.49, 637.18) mm, rotated rx -126.06 ry -5.23 rz 172.86 deg; joints [33.603, 114.274, -160.59, 72.301, 26.528, 52.723, 3120.904, 3490.151, 720.778]
  MoveL 182 to (1530.1, 797.35, 629.59) mm, rotated rx -125.49 ry -5.54 rz 172.29 deg; joints [33.55, 113.974, -160.59, 72.269, 27.436, 52.723, 3170.153, 3490.151, 727.159]
  MoveL 183 to (1571.43, 793.43, 622) mm, rotated rx -126.36 ry -6.17 rz 171.7 deg; joints [33.678, 113.974, -161.534, 73.024, 27.436, 52.723, 3225.026, 3481.37, 722.239]
  MoveL 184 to (1603.09, 790.02, 615.99) mm, rotated rx -125.07 ry -7.05 rz 170.09 deg; joints [33.678, 113.109, -161.582, 73.087, 29.648, 52.723, 3275.022, 3486.215, 722.239]
  MoveL 185 to (1632.65, 786.1, 609.97) mm, rotated rx -121.53 ry -6.97 rz 168.82 deg; joints [32.468, 113.109, -161.33, 72.481, 33.588, 52.723, 3301.948, 3486.215, 754.871]
  MoveL 186 to (1604.14, 786.62, 621.48) mm, rotated rx -118.75 ry -5.87 rz 169.45 deg; joints [31.246, 113.109, -159.904, 71.212, 35.486, 52.723, 3245.588, 3486.216, 774.116]
  Set speed (1000.0 mm/s)
  MoveL 187 to (1604.14, 786.62, 621.48) mm, rotated rx -118.75 ry -5.87 rz 169.45 deg; joints [31.246, 113.109, -159.904, 71.212, 35.486, 52.723, 3245.588, 3486.216, 774.116]
  MoveL 188 to (1625.03, 871.91, 669.33) mm, rotated rx -118.75 ry -5.87 rz 169.45 deg; joints [31.246, 113.109, -159.904, 71.212, 35.486, 52.723, 3266.48, 3571.502, 726.265]
  Set speed (1000.0 mm/s)
  MoveL 189 to (944.76, 961.41, 628.52) mm, rotated rx -102.53 ry -0.15 rz 179.33 deg; joints [22.48, 113.109, -152.046, 60.314, 43.621, 52.723, 2378.942, 3571.502, 957.472]
  MoveL 190 to (943.56, 863.8, 606.83) mm, rotated rx -102.53 ry -0.15 rz 179.33 deg; joints [22.48, 113.109, -152.046, 60.314, 43.621, 52.723, 2377.738, 3473.892, 979.167]
  MoveL 191 to (943.56, 863.8, 606.83) mm, rotated rx -102.53 ry -0.15 rz 179.33 deg; joints [22.48, 113.109, -152.046, 60.314, 43.621, 52.723, 2377.738, 3473.892, 979.167]
  Set speed (200.0 mm/s)
  MoveL 192 to (941.47, 865.37, 600.81) mm, rotated rx -103.3 ry -0.03 rz 179.89 deg; joints [22.48, 113.109, -152.046, 60.227, 42.743, 53.164, 2370.668, 3471.796, 979.259]
  MoveL 193 to (942.51, 867.72, 592.44) mm, rotated rx -104.82 ry 0.09 rz -179.67 deg; joints [22.635, 113.379, -152.046, 60.966, 41.175, 53.192, 2368.53, 3471.796, 979.256]
  MoveL 194 to (948.53, 871.13, 580.67) mm, rotated rx -104.47 ry 0.2 rz -179.23 deg; joints [22.461, 113.379, -151.846, 60.518, 41.165, 53.274, 2368.53, 3471.796, 995.471]
  MoveL 195 to (961.35, 877.14, 557.65) mm, rotated rx -101.65 ry 0.35 rz -178.31 deg; joints [21.918, 113.379, -151.344, 58.304, 42.654, 53.274, 2367.518, 3471.796, 1045.45]
  MoveL 196 to (968.94, 884.47, 522.07) mm, rotated rx -98.82 ry 0.38 rz -177.58 deg; joints [21.394, 113.036, -151.344, 55.674, 44.685, 53.957, 2366.085, 3471.796, 1100]
  MoveL 197 to (959.52, 887.08, 495.38) mm, rotated rx -96 ry 0.33 rz -176.86 deg; joints [21.363, 109.565, -151.344, 50.43, 48.362, 58.052, 2355.854, 3471.797, 1100]
  MoveL 198 to (949.84, 888.13, 477.07) mm, rotated rx -93.88 ry 0.21 rz -176.84 deg; joints [21.342, 107.078, -151.344, 47.67, 51.524, 60.107, 2351.553, 3471.796, 1100]
  MoveL 199 to (939.64, 888.39, 457.97) mm, rotated rx -92.71 ry 0.15 rz -176.83 deg; joints [21.429, 105.064, -151.344, 45.847, 53.719, 61.731, 2347.453, 3471.796, 1100]
  MoveL 200 to (929.69, 888.65, 437.83) mm, rotated rx -92 ry 0.11 rz -176.83 deg; joints [21.49, 103.237, -151.344, 44.523, 55.502, 63.165, 2343.762, 3470.933, 1100]
  MoveL 201 to (920.8, 888.65, 416.9) mm, rotated rx -90.71 ry 0.04 rz -176.82 deg; joints [21.49, 100.987, -151.344, 42.933, 58.101, 64.627, 2343.161, 3467.92, 1099.993]
  MoveL 202 to (912.69, 888.13, 394.4) mm, rotated rx -89.41 ry -0.04 rz -176.35 deg; joints [21.49, 98.6, -151.344, 40.968, 60.666, 66.288, 2341.199, 3461.341, 1100]
  MoveL 203 to (905.89, 887.61, 373.21) mm, rotated rx -88.94 ry -0.08 rz -175.41 deg; joints [21.49, 96.782, -151.344, 39.168, 62.052, 67.912, 2335.131, 3453.109, 1100]
  MoveL 204 to (900.66, 886.82, 356.2) mm, rotated rx -88.24 ry -0.14 rz -175.42 deg; joints [21.49, 94.919, -150.64, 38.552, 63.497, 68.439, 2335.131, 3450.131, 1100]
  MoveL 205 to (895.95, 886.04, 340.77) mm, rotated rx -88.24 ry -0.14 rz -175.42 deg; joints [21.49, 93.7, -150.334, 38.273, 64.212, 69.071, 2335.131, 3447.494, 1100]
  Set speed (1000.0 mm/s)
  MoveL 206 to (895.95, 886.04, 340.77) mm, rotated rx -88.24 ry -0.14 rz -175.42 deg; joints [21.49, 93.7, -150.334, 38.273, 64.212, 69.071, 2335.131, 3447.494, 1100]
  MoveL 207 to (887.95, 985.67, 337.69) mm, rotated rx -88.24 ry -0.14 rz -175.42 deg; joints [21.425, 93.472, -150.334, 38.273, 64.413, 69.196, 2328.017, 3545.651, 1100]
  Set speed (1000.0 mm/s)
  MoveL 208 to (853.38, 969.89, 348.17) mm, rotated rx -103.01 ry 7.43 rz -150.75 deg; joints [21.425, 93.472, -150.334, 9.922, 49.835, 97.581, 2115.612, 3359.096, 994.29]
  MoveL 209 to (903.53, 886.3, 325.86) mm, rotated rx -103.01 ry 7.43 rz -150.75 deg; joints [21.425, 93.472, -150.334, 9.922, 49.835, 97.581, 2165.763, 3275.508, 1016.606]
  MoveL 210 to (903.53, 886.3, 325.86) mm, rotated rx -103.01 ry 7.43 rz -150.75 deg; joints [21.425, 93.472, -150.334, 9.922, 49.835, 97.581, 2165.763, 3275.508, 1016.606]
  Set speed (200.0 mm/s)
  MoveL 211 to (914.52, 887.87, 345.22) mm, rotated rx -100.5 ry 6.57 rz -148.31 deg; joints [22.118, 93.472, -149.767, 6.474, 50.738, 97.381, 2165.763, 3275.326, 1016.606]
  MoveL 212 to (923.42, 888.65, 365.1) mm, rotated rx -102.16 ry 7.09 rz -150.22 deg; joints [21.962, 93.472, -149.766, 8.81, 49.725, 97.381, 2182.992, 3285.205, 984.925]
  MoveL 213 to (934.14, 889.44, 387.07) mm, rotated rx -103.41 ry 7.4 rz -151.62 deg; joints [21.92, 93.472, -149.767, 10.449, 48.952, 97.381, 2200.549, 3293.301, 953.912]
  MoveL 214 to (946.44, 890.22, 410.1) mm, rotated rx -105.74 ry 8.32 rz -152.83 deg; joints [21.683, 93.472, -149.758, 11.746, 47.568, 98.672, 2216.557, 3293.302, 915.548]
  MoveL 215 to (959.78, 890.48, 431.55) mm, rotated rx -108.87 ry 9.31 rz -154.67 deg; joints [21.399, 93.472, -149.758, 13.694, 45.669, 100.099, 2236.545, 3293.302, 872.978]
  MoveL 216 to (974.43, 890.75, 451.95) mm, rotated rx -110.73 ry 9.77 rz -155.85 deg; joints [21.224, 93.472, -149.758, 14.989, 44.51, 100.768, 2255.807, 3293.302, 839.728]
  MoveL 217 to (990.13, 890.48, 471.05) mm, rotated rx -114.55 ry 10.34 rz -158.54 deg; joints [20.905, 93.472, -149.758, 18.008, 42.046, 101.659, 2283.287, 3293.302, 793.397]
  MoveL 218 to (1011.58, 890.22, 492.77) mm, rotated rx -108.25 ry 10.08 rz -152.05 deg; joints [20.905, 93.472, -149.758, 10.729, 46.351, 102.075, 2270.138, 3267.055, 820.098]
  MoveL 219 to (1023.61, 888.13, 515.53) mm, rotated rx -113.08 ry 11.73 rz -154.49 deg; joints [20.905, 94.219, -149.758, 12.318, 42.718, 105.094, 2287.457, 3267.055, 776.725]
  Set speed (1000.0 mm/s)
  MoveL 220 to (1023.61, 888.13, 515.53) mm, rotated rx -113.08 ry 11.73 rz -154.49 deg; joints [20.905, 94.219, -149.758, 12.318, 42.718, 105.094, 2287.457, 3267.055, 776.725]
  MoveL 221 to (976.81, 967.73, 553.91) mm, rotated rx -113.08 ry 11.73 rz -154.49 deg; joints [20.905, 94.219, -149.758, 12.318, 42.718, 105.094, 2240.65, 3346.653, 738.343]

--- program FrameR_C (robot ABB IRB 1300-10/1.15) ---
  Smooth(1)
  Set speed (1000.0 mm/s)
  Set Ref.: FrameR
  Set Tool: Generic Paint Sprayer
  Show Generic Paint Sprayer
  MoveJ 1 to (-1567.41, -947.44, 561.3) mm, rotated rx 116.18 ry 8.07 rz 164.06 deg; joints [-18.613, 70.643, -160.975, 159.818, -72.367, 68.936, 14.365, 240.215, 405.979]
  MoveL 2 to (-1567.41, -947.44, 561.3) mm, rotated rx 116.18 ry 8.07 rz 164.06 deg; joints [-18.613, 70.643, -160.975, 159.818, -72.367, 68.936, 14.365, 240.215, 405.979]
  MoveL 3 to (-1536.8, -862.85, 517.62) mm, rotated rx 116.18 ry 8.07 rz 164.06 deg; joints [-18.613, 70.643, -160.975, 159.818, -72.367, 68.936, 44.975, 324.8, 449.664]
  MoveL 4 to (-1536.8, -862.85, 517.62) mm, rotated rx 116.18 ry 8.07 rz 164.06 deg; joints [-18.613, 70.643, -160.975, 159.818, -72.367, 68.936, 44.975, 324.8, 449.664]
  Set speed (200.0 mm/s)
  MoveL 5 to (-1511.42, -864.68, 530.96) mm, rotated rx 117.6 ry 7.57 rz 165.86 deg; joints [-18.613, 70.643, -160.975, 158.345, -70.921, 68.501, 83.279, 316.894, 423.259]
  MoveL 6 to (-1485.52, -866.25, 542.73) mm, rotated rx 119.49 ry 6.77 rz 168.23 deg; joints [-18.613, 70.643, -160.989, 156.392, -68.942, 68.006, 127.136, 308.433, 393.799]
  MoveL 7 to (-1458.84, -867.56, 552.68) mm, rotated rx 120.63 ry 6.22 rz 169.63 deg; joints [-18.608, 70.645, -160.989, 155.208, -67.701, 67.76, 164.896, 303.689, 373.04]
  MoveL 8 to (-1431.63, -868.61, 560.79) mm, rotated rx 121.87 ry 5.07 rz 171.91 deg; joints [-18.608, 70.645, -161.394, 153.058, -66.382, 67.76, 214.467, 295.937, 351.142]
  MoveL 9 to (-1403.9, -869.65, 567.06) mm, rotated rx 122.48 ry 4.46 rz 173.04 deg; joints [-18.608, 70.645, -161.65, 151.982, -65.747, 67.76, 254.1, 292.049, 337.984]
  MoveL 10 to (-1375.91, -870.7, 571.77) mm, rotated rx 122.85 ry 3.63 rz 174.4 deg; joints [-18.607, 70.645, -162.511, 150.654, -65.699, 67.76, 300.795, 287.554, 327.831]
  MoveL 11 to (-1347.65, -871.48, 574.39) mm, rotated rx 123.43 ry 2.18 rz 176.71 deg; joints [-18.607, 70.645, -163.965, 148.372, -65.568, 67.76, 361.589, 281.477, 316.442]
  MoveL 12 to (-1319.14, -872.53, 575.44) mm, rotated rx 123.01 ry 1.1 rz 178.31 deg; joints [-18.607, 70.645, -164.386, 146.346, -65.568, 68.646, 409.222, 272.173, 314.488]
  MoveL 13 to (-1290.62, -873.32, 574.39) mm, rotated rx 122.75 ry 0.03 rz 179.95 deg; joints [-18.607, 70.645, -164.966, 144.398, -65.568, 69.295, 458.433, 264.711, 313.88]
  MoveL 14 to (-1262.63, -874.1, 571.51) mm, rotated rx 121.5 ry -0.87 rz -178.58 deg; joints [-18.607, 70.645, -164.966, 142.218, -65.996, 70.794, 501.334, 252.628, 322.32]
  MoveL 15 to (-1234.64, -874.62, 567.06) mm, rotated rx 119.59 ry -1.16 rz -177.95 deg; joints [-18.607, 70.645, -164.966, 140.919, -67.366, 72.2, 535.411, 241.481, 339.756]
  MoveL 16 to (-1207.43, -875.41, 561.05) mm, rotated rx 117.47 ry -1.89 rz -176.36 deg; joints [-18.607, 70.645, -164.966, 138.54, -68.641, 74.029, 577.946, 226.627, 358.999]
  MoveL 17 to (-1181.01, -875.67, 553.72) mm, rotated rx 114.97 ry -2.36 rz -174.95 deg; joints [-18.607, 70.645, -164.966, 136.4, -70.403, 75.823, 617.522, 212.418, 383.818]
  MoveL 18 to (-1155.11, -876.19, 544.57) mm, rotated rx 113.17 ry -2.69 rz -173.75 deg; joints [-18.607, 70.645, -164.966, 134.745, -71.68, 77.07, 654.392, 202.078, 405.856]
  MoveL 19 to (-1130.25, -876.46, 534.1) mm, rotated rx 110.41 ry -2.6 rz -173.06 deg; joints [-18.607, 70.645, -164.966, 133.557, -74.022, 78.489, 684.783, 190.934, 438.633]
  MoveL 20 to (-1106.18, -876.46, 522.33) mm, rotated rx 107.69 ry -2.35 rz -172.66 deg; joints [-18.607, 70.645, -164.966, 132.771, -76.442, 79.73, 711.467, 182.061, 473.425]
  MoveL 21 to (-1082.9, -876.72, 508.72) mm, rotated rx 105 ry -2.28 rz -171.55 deg; joints [-18.607, 70.645, -164.966, 131.287, -78.713, 81.041, 744.285, 172.206, 509.473]
  MoveL 22 to (-1060.66, -876.46, 493.81) mm, rotated rx 102.34 ry -1.62 rz -172.64 deg; joints [-18.368, 70.645, -164.966, 131.892, -81.381, 81.898, 754.662, 172.209, 549.165]
  MoveL 23 to (-1048.89, -876.46, 484.92) mm, rotated rx 101.61 ry -1.74 rz -171.59 deg; joints [-18.368, 70.645, -164.966, 130.744, -81.892, 82.332, 775.999, 168.058, 563.788]
  Set speed (1000.0 mm/s)
  MoveL 24 to (-1048.89, -876.46, 484.92) mm, rotated rx 101.61 ry -1.74 rz -171.59 deg; joints [-18.368, 70.645, -164.966, 130.744, -81.892, 82.332, 775.999, 168.058, 563.788]
  MoveL 25 to (-1033.96, -973.27, 505.03) mm, rotated rx 101.61 ry -1.74 rz -171.59 deg; joints [-18.368, 70.645, -164.966, 130.744, -81.892, 82.332, 790.935, 71.246, 543.68]
  Set speed (1000.0 mm/s)
  MoveL 26 to (-1620.34, -905.96, 635.31) mm, rotated rx 95.09 ry -1.66 rz -161.98 deg; joints [-23.506, 70.645, -168.71, 125.797, -89.471, 82.332, 337.544, 71.246, 474.728]
  MoveL 27 to (-1651.39, -811.31, 626.45) mm, rotated rx 95.09 ry -1.66 rz -161.98 deg; joints [-23.507, 70.645, -168.71, 125.798, -89.471, 82.332, 306.493, 165.888, 483.588]
  MoveL 28 to (-1651.39, -811.31, 626.45) mm, rotated rx 95.09 ry -1.66 rz -161.98 deg; joints [-23.507, 70.645, -168.71, 125.798, -89.471, 82.332, 306.493, 165.888, 483.588]
  Set speed (200.0 mm/s)
  MoveL 29 to (-1645.89, -808.17, 640.32) mm, rotated rx 113.53 ry -8.08 rz -162.12 deg; joints [-23.507, 72.673, -168.71, 127.007, -69.184, 79.927, 306.494, 206.634, 309.416]
  MoveL 30 to (-1651.65, -799.02, 663.34) mm, rotated rx 121.42 ry -9.52 rz -164.85 deg; joints [-23.507, 72.673, -168.71, 130.57, -61.954, 76.902, 284.437, 252.951, 222.205]
  MoveL 31 to (-1666.56, -784.63, 693.42) mm, rotated rx 124.61 ry -9.92 rz -165.99 deg; joints [-23.507, 73.957, -168.71, 131.64, -58.294, 76.527, 250.715, 279.424, 178.795]
  MoveL 32 to (-1677.55, -774.95, 712.52) mm, rotated rx 126.3 ry -10.62 rz -165.92 deg; joints [-23.574, 73.957, -168.71, 131.661, -56.497, 76.164, 244.342, 297.996, 145.936]
  MoveL 33 to (-1683.83, -769.72, 722.72) mm, rotated rx 125.13 ry -10.25 rz -165.82 deg; joints [-23.558, 73.957, -169.107, 131.661, -57.93, 76.164, 239.386, 297.902, 145.355]
  MoveL 34 to (-1683.83, -769.72, 722.72) mm, rotated rx 171.16 ry 2.79 rz 179.57 deg; joints [-36.296, 73.957, -189.291, 194.827, -57.93, 27.33, 239.385, 619.77, 42.153]
  MoveL 35 to (-1643.8, -776.52, 722.72) mm, rotated rx 171.27 ry 13.42 rz 177.96 deg; joints [-36.914, 73.957, -189.291, 200.842, -67.394, 24.825, 197.215, 619.774, 96.315]
  MoveL 36 to (-1607.96, -779.4, 730.31) mm, rotated rx 167.94 ry 10.28 rz 177.82 deg; joints [-33.158, 73.957, -189.291, 194.194, -66.22, 26.961, 238.044, 614.627, 76.195]
  MoveL 37 to (-1574.47, -782.8, 735.54) mm, rotated rx 162.76 ry 12.18 rz 176.26 deg; joints [-33.158, 73.957, -186.255, 192.105, -66.997, 30.46, 238.043, 566.815, 81.388]
  Set speed (1000.0 mm/s)
  MoveL 38 to (-1574.47, -782.8, 735.54) mm, rotated rx 162.76 ry 12.18 rz 176.26 deg; joints [-33.158, 73.957, -186.255, 192.105, -66.997, 30.46, 238.043, 566.815, 81.388]
  MoveL 39 to (-1596.51, -811.05, 828.9) mm, rotated rx 162.76 ry 12.18 rz 176.26 deg; joints [-33.158, 75.195, -187.492, 192.105, -66.997, 30.46, 213.238, 536.755, 0.003]
  Set speed (1000.0 mm/s)
  MoveL 40 to (-1593.63, -878.91, 757.51) mm, rotated rx 98.12 ry 1.45 rz 169.97 deg; joints [-33.158, 75.195, -183.445, 163.358, -101.211, 79.486, 213.238, 138.256, 406.615]
  MoveL 41 to (-1576.04, -781.49, 743.39) mm, rotated rx 98.12 ry 1.45 rz 169.97 deg; joints [-33.158, 75.195, -183.445, 163.358, -101.211, 79.486, 230.829, 235.678, 420.735]
  MoveL 42 to (-1576.04, -781.49, 743.39) mm, rotated rx 98.12 ry 1.45 rz 169.97 deg; joints [-33.158, 75.195, -183.445, 163.358, -101.211, 79.486, 230.829, 235.678, 420.735]
  Set speed (200.0 mm/s)
  MoveL 43 to (-1574.47, -782.27, 739.73) mm, rotated rx 97.18 ry 1.28 rz 169.93 deg; joints [-33.158, 75.195, -183.201, 163.264, -101.701, 80.152, 230.829, 233.1, 431.046]
  MoveL 44 to (-1571.6, -783.32, 735.54) mm, rotated rx 102.36 ry 2.06 rz 170.68 deg; joints [-33.158, 75.729, -183.201, 163.488, -97.124, 76.98, 234.295, 233.103, 398.064]
  MoveL 45 to (-1568.19, -785.41, 730.05) mm, rotated rx 108.49 ry 2.67 rz 172.07 deg; joints [-33.158, 76.713, -183.201, 163.595, -91.261, 73.401, 239.31, 233.102, 362.103]
  MoveL 46 to (-1563.75, -789.08, 722.2) mm, rotated rx 111.32 ry 2.84 rz 172.75 deg; joints [-33.158, 76.962, -183.201, 163.705, -88.725, 71.728, 246.486, 233.102, 349.55]
  MoveL 47 to (-1557.21, -794.31, 711.74) mm, rotated rx 113.21 ry 2.87 rz 173.35 deg; joints [-33.158, 76.962, -183.201, 163.673, -87.145, 70.589, 257.356, 231.07, 345.118]
  MoveL 48 to (-1543.86, -806.08, 689.5) mm, rotated rx 112.74 ry 3 rz 172.89 deg; joints [-32.822, 76.962, -182.72, 163.673, -87.145, 70.89, 262.386, 220.973, 370.252]
  MoveL 49 to (-1538.37, -810.27, 681.65) mm, rotated rx 112.52 ry 3.31 rz 172.07 deg; joints [-32.75, 76.961, -182.72, 164.391, -87.566, 70.949, 260.5, 220.973, 381.211]
  MoveL 50 to (-1531.83, -814.19, 674.59) mm, rotated rx 113.2 ry 2.69 rz 173.74 deg; joints [-32.75, 76.961, -182.72, 162.867, -86.528, 70.657, 281.259, 210.637, 380.287]
  MoveL 51 to (-1524.51, -817.85, 668.31) mm, rotated rx 113.92 ry 2.93 rz 173.42 deg; joints [-32.75, 76.961, -182.72, 163.435, -86.107, 70.178, 285.413, 211.149, 381.936]
  MoveL 52 to (-1516.4, -821.25, 663.08) mm, rotated rx 112.76 ry 3.01 rz 172.86 deg; joints [-32.542, 76.961, -182.257, 163.435, -86.681, 70.937, 285.42, 206.557, 395.395]
  MoveL 53 to (-1507.76, -824.39, 658.89) mm, rotated rx 109.21 ry 2.91 rz 171.71 deg; joints [-32.402, 76.916, -182.257, 163.435, -89.666, 73.068, 285.419, 199.674, 427.279]
  MoveL 54 to (-1498.61, -826.75, 656.01) mm, rotated rx 109.9 ry 2.54 rz 173.03 deg; joints [-32.402, 76.916, -182.258, 162.277, -88.785, 72.69, 305.443, 192.437, 423.021]
  MoveL 55 to (-1489.19, -828.84, 654.18) mm, rotated rx 107.78 ry 2.44 rz 172.43 deg; joints [-32.365, 76.916, -181.423, 162.277, -89.745, 74.227, 305.447, 184.607, 439.56]
  MoveL 56 to (-1479.51, -830.41, 653.66) mm, rotated rx 108.96 ry 2.29 rz 173.36 deg; joints [-32.365, 76.916, -181.423, 161.636, -88.611, 73.537, 322.581, 181.509, 429.869]
  MoveL 57 to (-1428.23, -836.69, 652.87) mm, rotated rx 112.95 ry 1.82 rz 175.71 deg; joints [-32.365, 76.916, -181.424, 160.346, -84.86, 71.308, 393.108, 176.138, 396.691]
  MoveL 58 to (-1385.33, -840.88, 652.09) mm, rotated rx 113.89 ry 1.35 rz 176.95 deg; joints [-32.365, 76.916, -181.424, 159.328, -83.722, 70.904, 447.029, 169.407, 388.191]
  MoveL 59 to (-1341.9, -844.02, 651.57) mm, rotated rx 113.18 ry 1.15 rz 177.32 deg; joints [-32.365, 76.916, -181.269, 158.734, -84.013, 71.415, 492.999, 161.611, 393.106]
  MoveL 60 to (-1314.69, -845.58, 651.04) mm, rotated rx 113.65 ry 1.17 rz 177.34 deg; joints [-32.249, 77.105, -181.269, 158.734, -83.449, 71.189, 518.198, 161.611, 391.36]
  MoveL 61 to (-1305.01, -845.58, 652.35) mm, rotated rx 113.89 ry 1.18 rz 177.34 deg; joints [-32.235, 77.284, -181.269, 158.773, -83.092, 71.116, 526.446, 161.611, 389.548]
  MoveL 62 to (-1296.12, -844.28, 656.27) mm, rotated rx 112.25 ry 0.44 rz 178.92 deg; joints [-32.235, 77.284, -181.226, 156.661, -83.843, 72.256, 549.803, 150.421, 395.544]
  MoveL 63 to (-1288.27, -842.18, 662.29) mm, rotated rx 109.89 ry -0.2 rz -179.46 deg; joints [-32.235, 77.284, -181.225, 154.389, -85.281, 73.661, 572.589, 138.737, 405.907]
  MoveL 64 to (-1282.25, -839.04, 669.88) mm, rotated rx 113.65 ry 0.48 rz 178.91 deg; joints [-32.235, 77.286, -181.23, 157.059, -82.712, 71.482, 563.484, 160.403, 371.001]
  MoveL 65 to (-1278.85, -835.12, 679.03) mm, rotated rx 113.65 ry 0.13 rz 179.7 deg; joints [-32.317, 77.286, -181.23, 156.309, -82.452, 71.61, 574.687, 160.404, 360.488]
  MoveL 66 to (-1277.54, -830.93, 688.71) mm, rotated rx 113.66 ry 0.65 rz 178.52 deg; joints [-32.317, 77.71, -181.23, 157.531, -82.452, 71.603, 561.67, 167.436, 355.878]
  MoveL 67 to (-1279.11, -826.49, 698.39) mm, rotated rx 113.19 ry 1.66 rz 176.12 deg; joints [-32.317, 77.959, -181.23, 159.893, -83.38, 71.634, 536.353, 179.707, 355.876]
  MoveL 68 to (-1282.51, -822.82, 706.5) mm, rotated rx 112.01 ry 1.43 rz 176.46 deg; joints [-32.317, 77.951, -181.23, 159.203, -84.202, 72.371, 536.352, 177.924, 356.114]
  MoveL 69 to (-1287.22, -818.9, 715.4) mm, rotated rx 109.18 ry 1.43 rz 175.91 deg; joints [-32.485, 77.234, -181.23, 159.196, -87.271, 73.747, 533.82, 177.924, 364.649]
  MoveL 70 to (-1291.67, -816.02, 722.99) mm, rotated rx 105.18 ry 1.04 rz 176.17 deg; joints [-32.485, 77.049, -181.23, 157.979, -90.559, 75.959, 533.82, 170.277, 387.037]
  MoveL 71 to (-1294.81, -814.45, 728.74) mm, rotated rx 100.47 ry 0.65 rz 176.47 deg; joints [-32.485, 77.049, -181.224, 156.739, -94.298, 78.535, 533.825, 161.41, 419.179]
  MoveL 72 to (-1297.16, -813.67, 732.67) mm, rotated rx 97.77 ry 0.62 rz 175.5 deg; joints [-32.485, 77.049, -181.224, 157.267, -96.675, 80.1, 523.529, 162.939, 438.079]
  MoveL 73 to (-1298.99, -813.14, 736.07) mm, rotated rx 89.91 ry -0.01 rz 175.41 deg; joints [-32.485, 76.771, -181.224, 156.398, -103.36, 84.313, 523.529, 160.679, 497.487]
  Set speed (1000.0 mm/s)
  MoveL 74 to (-1298.99, -813.14, 736.07) mm, rotated rx 89.91 ry -0.01 rz 175.41 deg; joints [-32.485, 76.771, -181.224, 156.398, -103.36, 84.313, 523.529, 160.679, 497.487]
  MoveL 75 to (-1306.99, -912.82, 735.92) mm, rotated rx 89.91 ry -0.01 rz 175.41 deg; joints [-32.485, 76.771, -181.224, 156.398, -103.36, 84.313, 515.53, 61, 497.634]
  Set speed (1000.0 mm/s)
  MoveL 76 to (-1277.26, -812.46, 899.51) mm, rotated rx 130.43 ry 1.94 rz 177.73 deg; joints [-32.485, 82.485, -181.224, 164.314, -65.405, 62.278, 515.529, 241.607, 65.66]
  MoveL 77 to (-1272.05, -736.49, 834.7) mm, rotated rx 130.43 ry 1.94 rz 177.73 deg; joints [-32.485, 82.485, -181.224, 164.314, -65.405, 62.278, 520.743, 317.58, 130.474]
  MoveL 78 to (-1272.05, -736.49, 834.7) mm, rotated rx 130.43 ry 1.94 rz 177.73 deg; joints [-32.485, 82.485, -181.224, 164.314, -65.405, 62.278, 520.743, 317.58, 130.474]
  Set speed (200.0 mm/s)
  MoveL 79 to (-1313.64, -732.57, 835.74) mm, rotated rx 131.13 ry 1.86 rz 177.87 deg; joints [-32.486, 82.485, -181.225, 164.465, -64.816, 61.836, 480.451, 324.806, 124.566]
  MoveL 80 to (-1348.7, -729.17, 836.53) mm, rotated rx 131.51 ry 2.46 rz 177.23 deg; joints [-32.486, 82.585, -181.206, 165.473, -64.817, 61.212, 437.294, 332.811, 124.566]
  MoveL 81 to (-1370.15, -726.81, 837.05) mm, rotated rx 131.03 ry 2.25 rz 177.41 deg; joints [-32.486, 82.375, -181.206, 165.02, -65.244, 61.624, 419.632, 332.534, 124.566]
  MoveL 82 to (-1401.81, -723.67, 837.57) mm, rotated rx 132.04 ry 2.5 rz 177.23 deg; joints [-32.486, 82.375, -181.206, 165.762, -64.645, 60.747, 385.483, 342.305, 118.589]
  MoveL 83 to (-1441.84, -719.23, 838.1) mm, rotated rx 133.18 ry 2.93 rz 176.89 deg; joints [-32.49, 82.375, -181.783, 166.881, -64.645, 59.499, 344.476, 357.293, 113.753]
  MoveL 84 to (-1485.26, -713.73, 838.88) mm, rotated rx 133.65 ry 3 rz 176.86 deg; joints [-32.492, 82.375, -182.089, 167.201, -64.645, 59.035, 302.34, 366.865, 110.952]
  MoveL 85 to (-1528.43, -707.71, 839.4) mm, rotated rx 134.21 ry 4.21 rz 175.68 deg; joints [-32.492, 82.375, -181.644, 169.049, -64.645, 57.959, 242.645, 380.514, 111.34]
  MoveL 86 to (-1562.18, -702.74, 839.67) mm, rotated rx 135.2 ry 4.73 rz 175.31 deg; joints [-32.493, 82.375, -181.868, 170.148, -64.51, 56.845, 205.151, 394.369, 107.799]
  MoveL 87 to (-1610.05, -694.63, 839.67) mm, rotated rx 135.22 ry 5.08 rz 174.98 deg; joints [-32.493, 82.375, -181.638, 170.602, -64.511, 56.652, 152, 403.576, 108.755]
  MoveL 88 to (-1652.17, -686.26, 839.67) mm, rotated rx 135.73 ry 5.47 rz 174.69 deg; joints [-32.493, 82.375, -181.727, 171.316, -64.511, 56.005, 106.555, 417.077, 107.647]
  MoveL 89 to (-1691.68, -677.63, 839.67) mm, rotated rx 136.03 ry 5.85 rz 174.38 deg; joints [-32.493, 82.383, -181.727, 171.926, -64.56, 55.539, 63.117, 429.319, 107.647]
  MoveL 90 to (-1724.9, -670.56, 838.1) mm, rotated rx 136.82 ry 6.43 rz 174 deg; joints [-32.493, 82.383, -181.876, 172.973, -64.56, 54.549, 25.38, 444.226, 107.518]
  MoveL 91 to (-1758.39, -661.41, 836.26) mm, rotated rx 135.23 ry 8 rz 172.14 deg; joints [-34.724, 80.46, -181.876, 176.549, -68.763, 55.099, 0.002, 444.226, 110.987]
  Set speed (1000.0 mm/s)
  MoveL 92 to (-1758.39, -661.41, 836.26) mm, rotated rx 135.23 ry 8 rz 172.14 deg; joints [-34.724, 80.46, -181.876, 176.549, -68.763, 55.099, 0.002, 444.226, 110.987]
  MoveL 93 to (-1777.81, -729.83, 906.56) mm, rotated rx 135.23 ry 8 rz 172.14 deg; joints [-34.724, 80.46, -185.22, 176.62, -72.101, 54.888, 0, 389.269, 48.578]
  Set speed (1000.0 mm/s)
  MoveL 94 to (892.89, -973.97, 160.56) mm, rotated rx 74.09 ry -79.65 rz -165.04 deg; joints [-50.625, 101.986, -183.176, 143.958, -56.047, 174.635, 2943.702, -296.83, 1100]
  MoveL 95 to (894.12, -874.1, 165.49) mm, rotated rx 74.09 ry -79.65 rz -165.04 deg; joints [-50.625, 102.249, -183.176, 143.853, -55.834, 174.822, 2944.041, -198.044, 1097.78]
  MoveL 96 to (894.12, -874.1, 165.49) mm, rotated rx 74.09 ry -79.65 rz -165.04 deg; joints [-50.625, 102.249, -183.176, 143.853, -55.834, 174.822, 2944.041, -198.044, 1097.78]
  Set speed (200.0 mm/s)
  MoveL 97 to (897.25, -874.89, 176.21) mm, rotated rx 65.87 ry -79.15 rz -157.31 deg; joints [-50.572, 102.13, -183.176, 144.306, -57.481, 174.822, 2944.041, -202.933, 1099.813]
  MoveL 98 to (899.87, -876.46, 192.17) mm, rotated rx 61.84 ry -78.73 rz -152.65 deg; joints [-50.572, 102.13, -183.176, 143.646, -58.425, 174.912, 2952.705, -207.84, 1091.736]
  MoveL 99 to (903.01, -878.29, 209.44) mm, rotated rx 62.04 ry -78.65 rz -151.92 deg; joints [-50.572, 102.13, -183.176, 142.694, -58.517, 174.948, 2963.908, -210.297, 1074.532]
  MoveL 100 to (906.93, -880.12, 229.58) mm, rotated rx 62.24 ry -78.57 rz -151.18 deg; joints [-50.572, 102.13, -183.176, 141.745, -58.61, 174.982, 2975.895, -212.626, 1054.448]
  MoveL 101 to (912.69, -881.95, 251.82) mm, rotated rx 63.48 ry -78.61 rz -151.46 deg; joints [-50.572, 102.13, -183.22, 140.789, -58.506, 174.982, 2989.943, -213.842, 1030.144]
  MoveL 102 to (920.28, -883.78, 275.36) mm, rotated rx 64.54 ry -78.72 rz -152.5 deg; joints [-50.571, 102.13, -183.221, 140.765, -58.272, 174.982, 2997.54, -214.928, 1004.496]
  MoveL 103 to (929.69, -885.35, 299.69) mm, rotated rx 65.62 ry -78.83 rz -153.56 deg; joints [-50.545, 102.13, -183.227, 140.714, -58.045, 174.982, 3006.729, -215.496, 978.065]
  MoveL 104 to (940.68, -886.66, 324.29) mm, rotated rx 66.79 ry -78.9 rz -154.23 deg; joints [-50.519, 102.13, -183.265, 140.199, -57.891, 174.982, 3021.693, -215.76, 951.388]
  MoveL 105 to (953.5, -887.97, 348.36) mm, rotated rx 85.13 ry -19.62 rz -174.48 deg; joints [0, 44.016, -168.118, 113.546, -98.533, 78.32, 3060.514, 351.718, 637.921]
  MoveL 106 to (968.15, -889.01, 371.64) mm, rotated rx 85.13 ry -19.62 rz -174.48 deg; joints [0, 44.016, -168.118, 113.546, -98.533, 78.32, 3075.164, 350.671, 614.638]
  MoveL 107 to (984.11, -889.8, 393.88) mm, rotated rx 84.63 ry -19.58 rz -174.31 deg; joints [0, 44.835, -168.118, 113.424, -98.568, 79.239, 3080.491, 349.61, 598.511]
  MoveL 108 to (1001.38, -890.32, 415.07) mm, rotated rx 85.13 ry -19.62 rz -174.48 deg; joints [0.001, 44.853, -168.118, 113.658, -98.197, 79.096, 3097.541, 349.369, 573.162]
  MoveL 109 to (1020.21, -890.58, 435.21) mm, rotated rx 84.63 ry -19.58 rz -174.31 deg; joints [0.001, 45.265, -168.118, 113.481, -98.396, 79.637, 3111.032, 348.831, 558.239]
  MoveL 110 to (1040.1, -890.84, 453.79) mm, rotated rx 84.38 ry -19.55 rz -174.23 deg; joints [0.001, 45.523, -168.118, 113.402, -98.476, 79.957, 3127.571, 348.445, 542.424]
  MoveL 111 to (1066.78, -890.84, 475.24) mm, rotated rx 84.63 ry -19.58 rz -174.31 deg; joints [0.001, 45.532, -168.118, 113.517, -98.289, 79.885, 3154.15, 348.57, 518.893]
  MoveL 112 to (1095.03, -890.58, 494.6) mm, rotated rx 85.13 ry -19.62 rz -174.48 deg; joints [0.001, 45.549, -168.118, 113.748, -97.917, 79.739, 3182.208, 349.108, 495.375]
  MoveL 113 to (1124.86, -890.06, 511.6) mm, rotated rx 85.38 ry -19.72 rz -175.5 deg; joints [0.001, 45.558, -168.118, 114.693, -98.158, 79.939, 3203.662, 352.782, 476.029]
  MoveL 114 to (1155.99, -889.54, 525.99) mm, rotated rx 85.88 ry -19.72 rz -175.19 deg; joints [0, 45.573, -168.118, 114.51, -97.577, 79.649, 3238.754, 352.115, 457.625]
  MoveL 115 to (1181.63, -888.75, 535.67) mm, rotated rx 86.12 ry -19.77 rz -175.75 deg; joints [0, 45.582, -168.118, 115.04, -97.607, 79.708, 3260.15, 354.598, 445.767]
  MoveL 116 to (1207.79, -887.97, 543.52) mm, rotated rx 86.62 ry -19.83 rz -176.38 deg; joints [0, 45.6, -168.118, 115.686, -97.454, 79.686, 3281.974, 357.321, 433.7]
  MoveL 117 to (1234.47, -887.18, 549.8) mm, rotated rx 86.87 ry -19.87 rz -176.94 deg; joints [0, 45.613, -168.118, 116.215, -97.485, 79.743, 3304.394, 359.899, 425.291]
  MoveL 118 to (1261.68, -886.4, 554.25) mm, rotated rx 87.62 ry -19.89 rz -176.72 deg; joints [0, 45.625, -168.118, 116.15, -96.728, 79.358, 3335.564, 359.768, 414.744]
  MoveL 119 to (1288.89, -885.35, 556.86) mm, rotated rx 88.12 ry -19.93 rz -177.36 deg; joints [0, 45.643, -168.118, 116.795, -96.582, 79.323, 3358.44, 362.895, 407.98]
  MoveL 120 to (1316.36, -884.57, 557.91) mm, rotated rx 88.12 ry -19.96 rz -178.3 deg; joints [0.004, 45.662, -168.118, 117.618, -97.006, 79.598, 3377.48, 366.981, 406.875]
  MoveL 121 to (1343.57, -883.78, 556.86) mm, rotated rx 88.12 ry -19.96 rz -178.3 deg; joints [0.004, 45.662, -168.118, 117.618, -97.006, 79.598, 3404.688, 367.766, 407.922]
  MoveL 122 to (1371.04, -883, 554.25) mm, rotated rx 87.87 ry -19.95 rz -178.21 deg; joints [-0.098, 45.662, -168.118, 117.592, -97.231, 79.716, 3432.156, 367.766, 412.586]
  MoveL 123 to (1398.24, -882.21, 549.8) mm, rotated rx 88.12 ry -19.96 rz -178.3 deg; joints [-0.098, 45.668, -168.118, 117.708, -97.052, 79.628, 3459.294, 368.802, 415]
  MoveL 124 to (1425.45, -881.43, 543.52) mm, rotated rx 88.87 ry -19.98 rz -178.56 deg; joints [-0.098, 45.682, -168.118, 118.055, -96.518, 79.362, 3486.317, 370.389, 415.176]
  MoveL 125 to (1452.4, -880.64, 535.67) mm, rotated rx 88.87 ry -19.98 rz -178.56 deg; joints [-0.098, 45.682, -168.118, 118.055, -96.518, 79.362, 3513.264, 371.174, 423.025]
  Set speed (1000.0 mm/s)
  MoveL 126 to (1452.4, -880.64, 535.67) mm, rotated rx 88.87 ry -19.98 rz -178.56 deg; joints [-0.098, 45.682, -168.118, 118.055, -96.518, 79.362, 3513.264, 371.174, 423.025]
  MoveL 127 to (1454.25, -980.61, 533.82) mm, rotated rx 88.87 ry -19.98 rz -178.56 deg; joints [-0.098, 45.682, -168.118, 118.055, -96.518, 79.362, 3515.111, 271.208, 424.873]
  Set speed (1000.0 mm/s)
  MoveL 128 to (1533.99, -926.46, 631.09) mm, rotated rx 138.74 ry -6.11 rz -174.67 deg; joints [-9.541, 61.146, -158.442, 135.819, -50.553, 59.636, 3391.215, 390.14, 48.578]
  MoveL 129 to (1519.9, -861.54, 556.34) mm, rotated rx 138.74 ry -6.11 rz -174.67 deg; joints [-9.541, 61.146, -158.442, 135.819, -50.553, 59.636, 3377.12, 455.057, 123.326]
  MoveL 130 to (1519.9, -861.54, 556.34) mm, rotated rx 138.74 ry -6.11 rz -174.67 deg; joints [-9.541, 61.146, -158.442, 135.819, -50.553, 59.636, 3377.12, 455.057, 123.326]
  Set speed (200.0 mm/s)
  MoveL 131 to (1489.29, -872.53, 551.89) mm, rotated rx 138.33 ry -11.97 rz -169.54 deg; joints [-9.406, 61.146, -158.442, 126.772, -46.624, 65.411, 3417.685, 437.6, 113.159]
  MoveL 132 to (1461.56, -873.05, 561.57) mm, rotated rx 139.84 ry -10.86 rz -170.96 deg; joints [-9.406, 61.146, -158.442, 129.677, -46.276, 63.079, 3373.678, 447.966, 98.005]
  MoveL 133 to (1433.04, -873.58, 569.68) mm, rotated rx 141.66 ry -9.37 rz -172.66 deg; joints [-9.406, 61.146, -158.442, 133.371, -46.012, 60.06, 3324.622, 461.468, 84.178]
  MoveL 134 to (1404.52, -874.36, 576.22) mm, rotated rx 143.33 ry -7.53 rz -174.43 deg; joints [-9.406, 61.146, -158.442, 137.332, -46.181, 56.838, 3272.974, 474.662, 74.367]
  MoveL 135 to (1375.22, -875.15, 580.67) mm, rotated rx 143.54 ry -5.51 rz -175.94 deg; joints [-9.406, 61.073, -158.442, 140.257, -47.619, 54.789, 3221.713, 478.344, 74.674]
  MoveL 136 to (1345.92, -875.93, 583.81) mm, rotated rx 143.06 ry -3.49 rz -177.38 deg; joints [-9.406, 61.217, -158.628, 142.541, -49.547, 53.504, 3169.819, 477.803, 82.221]
  MoveL 137 to (1316.1, -876.98, 585.12) mm, rotated rx 142.32 ry -2.18 rz -178.32 deg; joints [-9.406, 61.43, -158.905, 143.697, -51.125, 53.088, 3125.253, 474.44, 91.484]
  MoveL 138 to (1286.01, -877.76, 585.38) mm, rotated rx 140.67 ry -0.69 rz -179.43 deg; joints [-9.406, 61.887, -159.499, 144.523, -53.535, 53.312, 3077.773, 466.28, 109.947]
  MoveL 139 to (1255.14, -878.55, 584.07) mm, rotated rx 137.84 ry 0.78 rz 179.29 deg; joints [-9.406, 62.612, -160.443, 144.766, -56.841, 54.489, 3028.427, 451.799, 139.793]
  MoveL 140 to (1223.49, -879.07, 581.45) mm, rotated rx 134.73 ry 1.74 rz 178.25 deg; joints [-9.406, 63.328, -161.381, 144.461, -59.978, 56.161, 2983.148, 436.266, 171.527]
  MoveL 141 to (1190.26, -879.59, 578.05) mm, rotated rx 133.24 ry 1.97 rz 177.91 deg; joints [-9.406, 63.653, -161.807, 144.091, -61.33, 57.095, 2945.816, 428.197, 188.24]
  MoveL 142 to (1155.47, -879.59, 573.87) mm, rotated rx 131.24 ry 2.37 rz 177.3 deg; joints [-9.406, 64.059, -162.341, 143.811, -63.215, 58.243, 2904.186, 419.258, 210.694]
  MoveL 143 to (1117.01, -879.07, 569.16) mm, rotated rx 126.69 ry 2.59 rz 176.53 deg; joints [-9.406, 64.918, -163.475, 142.508, -67.052, 61.172, 2857.854, 398.451, 254.993]
  MoveL 144 to (1084.05, -880.38, 560) mm, rotated rx 121.8 ry 2.47 rz 176.03 deg; joints [-9.406, 65.478, -164.218, 140.911, -70.931, 64.405, 2821.001, 375.562, 303.776]
  MoveL 145 to (1052.39, -880.9, 553.98) mm, rotated rx 120.88 ry 0.65 rz 178.91 deg; joints [-9.834, 65.478, -164.218, 137.662, -70.306, 66.212, 2818.641, 353.715, 309.094]
  MoveL 146 to (1009.23, -879.33, 553.98) mm, rotated rx 119.04 ry 0.4 rz 179.27 deg; joints [-10.314, 65.479, -164.219, 137.039, -71.636, 67.57, 2780.014, 341.197, 321.813]
  Set speed (1000.0 mm/s)
  MoveL 147 to (1009.23, -879.33, 553.98) mm, rotated rx 119.04 ry 0.4 rz 179.27 deg; joints [-10.314, 65.479, -164.219, 137.039, -71.636, 67.57, 2780.014, 341.197, 321.813]
  MoveL 148 to (1007.78, -966.75, 602.53) mm, rotated rx 119.04 ry 0.4 rz 179.27 deg; joints [-10.314, 65.479, -164.219, 137.039, -71.636, 67.57, 2778.565, 253.784, 273.265]
  Set speed (1000.0 mm/s)
  MoveL 149 to (873.5, -880.28, 780.09) mm, rotated rx 138.11 ry -2.37 rz -177.88 deg; joints [-10.314, 69.754, -169.974, 142.569, -56.185, 54.961, 2673.473, 430.431, 0]
  MoveL 150 to (867.95, -813.67, 705.72) mm, rotated rx 138.11 ry -2.37 rz -177.88 deg; joints [-10.314, 69.754, -169.974, 142.569, -56.185, 54.961, 2667.932, 497.048, 74.374]
  MoveL 151 to (867.95, -813.67, 705.72) mm, rotated rx 138.11 ry -2.37 rz -177.88 deg; joints [-10.314, 69.754, -169.974, 142.569, -56.185, 54.961, 2667.932, 497.048, 74.374]
  Set speed (200.0 mm/s)
  MoveL 152 to (904.84, -813.67, 702.84) mm, rotated rx 138.4 ry -2.86 rz -177.46 deg; joints [-10.348, 69.754, -169.974, 142.156, -55.592, 55.078, 2710.558, 497.291, 73.781]
  MoveL 153 to (941.47, -813.41, 700.23) mm, rotated rx 139.78 ry -3.56 rz -176.99 deg; joints [-10.348, 69.694, -169.893, 142.201, -54.052, 54.45, 2754.696, 505.196, 65.514]
  MoveL 154 to (978.09, -813.14, 697.35) mm, rotated rx 140.31 ry -3.04 rz -177.48 deg; joints [-10.213, 69.694, -169.893, 143.129, -54.093, 53.594, 2784.707, 511.736, 67.35]
  MoveL 155 to (1014.72, -812.62, 694.47) mm, rotated rx 138.88 ry -3.15 rz -177.25 deg; joints [-10.213, 69.694, -169.893, 141.972, -54.989, 54.887, 2823.471, 502.14, 77.761]
  MoveL 156 to (1051.87, -812.1, 691.59) mm, rotated rx 137.92 ry -3.25 rz -177.07 deg; joints [-10.214, 69.694, -169.893, 141.188, -55.584, 55.745, 2862.315, 495.937, 85.751]
  MoveL 157 to (1090.33, -811.58, 688.45) mm, rotated rx 140.78 ry -3.42 rz -177.21 deg; joints [-10.214, 69.645, -169.825, 142.984, -53.446, 53.474, 2901.1, 515.702, 71.782]
  MoveL 158 to (1131.14, -810.79, 684.79) mm, rotated rx 141.73 ry -3.41 rz -177.31 deg; joints [-10.214, 69.629, -169.804, 143.689, -52.802, 52.645, 2941.325, 523.172, 70.224]
  MoveL 159 to (1175.09, -810.01, 680.6) mm, rotated rx 141.49 ry -3.86 rz -176.93 deg; joints [-10.214, 69.629, -169.804, 142.952, -52.605, 53.185, 2990.491, 521.26, 74.11]
  MoveL 160 to (1220.35, -808.96, 676.16) mm, rotated rx 141.93 ry -4.58 rz -176.42 deg; joints [-10.239, 69.647, -169.804, 142.399, -51.718, 53.352, 3043.49, 523.666, 73.879]
  MoveL 161 to (1265.35, -807.91, 671.45) mm, rotated rx 142.71 ry -3.96 rz -176.99 deg; joints [-10.076, 69.647, -169.803, 143.629, -51.673, 52.164, 3080.695, 533.169, 76.64]
  MoveL 162 to (1308.25, -806.6, 666.74) mm, rotated rx 142.43 ry -3.78 rz -177.1 deg; joints [-10.029, 69.733, -169.803, 143.556, -51.931, 52.336, 3120.743, 533.169, 84.07]
  MoveL 163 to (1347.49, -805.3, 662.29) mm, rotated rx 142.24 ry -4.83 rz -176.27 deg; joints [-10.206, 69.7, -169.758, 142.247, -51.221, 53.337, 3172.343, 529.258, 85.549]
  MoveL 164 to (1385.43, -803.73, 657.84) mm, rotated rx 141.75 ry -6.36 rz -175.01 deg; joints [-10.206, 69.7, -169.758, 139.926, -50.344, 54.95, 3228.058, 524.713, 87.591]
  MoveL 165 to (1429.12, -801.37, 651.83) mm, rotated rx 140.48 ry -6.48 rz -174.69 deg; joints [-10.206, 69.7, -169.758, 138.77, -51.128, 56.142, 3274.416, 517.767, 100.02]
  MoveL 166 to (1480.65, -797.97, 643.98) mm, rotated rx 140.88 ry -6.94 rz -174.39 deg; joints [-10.551, 69.337, -169.263, 138.71, -50.428, 56.337, 3331.85, 520.017, 100.585]
  MoveL 167 to (1525.91, -794.57, 636.39) mm, rotated rx 143.15 ry -7.95 rz -174.08 deg; joints [-10.551, 69.344, -169.263, 139.263, -48.057, 55.155, 3386.01, 538.846, 93.227]
  MoveL 168 to (1570.39, -790.38, 628.28) mm, rotated rx 142.96 ry -9.33 rz -173.02 deg; joints [-10.712, 69.33, -169.245, 137.427, -47.121, 56.529, 3446.772, 538.846, 98.189]
  MoveL 169 to (1604.14, -786.72, 621.48) mm, rotated rx 141.05 ry -10.48 rz -171.64 deg; joints [-10.712, 69.329, -169.243, 134.243, -47.573, 59.2, 3496.639, 527.838, 111.781]
  MoveL 170 to (1635.01, -782.8, 614.94) mm, rotated rx 141.92 ry -11.12 rz -171.41 deg; joints [-10.712, 69.3, -169.204, 134.121, -46.464, 59.025, 3533.455, 537.973, 111.775]
  MoveL 171 to (1664.04, -778.61, 608.4) mm, rotated rx 141.82 ry -12.17 rz -170.59 deg; joints [-11.054, 69.025, -168.829, 132.808, -45.717, 60.235, 3575.747, 537.973, 113.449]
  MoveL 172 to (1691.25, -774.16, 601.34) mm, rotated rx 142.72 ry -13.83 rz -169.68 deg; joints [-11.054, 69.024, -168.829, 131.288, -43.831, 61.04, 3620.345, 549.538, 112.01]
  MoveL 173 to (1717.15, -769.46, 594.01) mm, rotated rx 144.18 ry -14.24 rz -169.93 deg; joints [-11.054, 69.024, -168.829, 132.075, -42.496, 60.144, 3647.995, 565.322, 111.216]
  MoveL 174 to (1741.48, -764.22, 585.9) mm, rotated rx 143.22 ry -16.98 rz -167.69 deg; joints [-11.113, 69.024, -168.829, 127.258, -41.194, 63.853, 3705.229, 565.239, 118.706]
  MoveL 175 to (1763.46, -759.25, 577.79) mm, rotated rx 147.1 ry -20.86 rz -167.03 deg; joints [-11.113, 69.024, -168.829, 125.179, -35.697, 64.914, 3760.726, 604.805, 103.148]
  MoveL 176 to (1782.03, -754.81, 570.47) mm, rotated rx 149.6 ry -22.53 rz -167.33 deg; joints [-11.113, 69.024, -168.828, 125.124, -32.775, 64.732, 3791.331, 631.104, 98.349]
  MoveL 177 to (1797.47, -750.88, 563.66) mm, rotated rx 149.1 ry -22.89 rz -166.9 deg; joints [-11.207, 68.767, -168.479, 123.926, -32.856, 65.888, 3812.138, 631.104, 104.311]
  MoveL 178 to (1809.5, -747.74, 557.91) mm, rotated rx 149.34 ry -27.13 rz -164.88 deg; joints [-11.369, 68.485, -168.097, 116.582, -30.027, 72.314, 3867.977, 644.455, 104.311]
  MoveL 179 to (1819.44, -745.39, 552.94) mm, rotated rx 152.47 ry -25.62 rz -167.3 deg; joints [-11.369, 69.123, -168.963, 123.151, -28.77, 66.476, 3854.856, 665.831, 104.31]
  MoveL 180 to (1827.81, -743.03, 548.23) mm, rotated rx 155.32 ry -27.01 rz -168.21 deg; joints [-11.369, 69.123, -168.963, 123.836, -25.853, 65.81, 3871.651, 692.676, 99.167]
  Set speed (1000.0 mm/s)
  MoveL 181 to (1827.81, -743.03, 548.23) mm, rotated rx 155.32 ry -27.01 rz -168.21 deg; joints [-11.369, 69.123, -168.963, 123.836, -25.853, 65.81, 3871.651, 692.676, 99.167]
  MoveL 182 to (1876.74, -775.47, 629.18) mm, rotated rx 155.32 ry -27.01 rz -168.21 deg; joints [-11.369, 69.123, -168.963, 123.836, -25.853, 65.81, 3920.576, 660.235, 18.211]
  Set speed (1000.0 mm/s)
  MoveL 183 to (883.17, -844.02, 851.21) mm, rotated rx 124.16 ry -6.87 rz -170 deg; joints [-11.369, 72, -172.918, 127.917, -63.476, 67.716, 2763.544, 357.619, 25.596]
  MoveL 184 to (862.2, -763.7, 795.45) mm, rotated rx 124.16 ry -6.87 rz -170 deg; joints [-11.369, 71.999, -172.918, 127.917, -63.476, 67.715, 2742.569, 437.942, 81.346]
  MoveL 185 to (862.2, -763.7, 795.45) mm, rotated rx 124.16 ry -6.87 rz -170 deg; joints [-11.369, 71.999, -172.918, 127.917, -63.476, 67.715, 2742.569, 437.942, 81.346]
  Set speed (200.0 mm/s)
  MoveL 186 to (834.21, -757.94, 813.24) mm, rotated rx 125.41 ry -7.49 rz -169.6 deg; joints [-11.997, 71.344, -172.918, 128.596, -62.551, 66.897, 2728.773, 444.882, 47.939]
  MoveL 187 to (805.69, -752.19, 831.29) mm, rotated rx 128.43 ry -8.31 rz -169.68 deg; joints [-12.476, 70.429, -172.918, 130.342, -60.33, 64.815, 2714.571, 464.902, 0.024]
  MoveL 188 to (775.87, -745.91, 849.87) mm, rotated rx 128.95 ry -7.87 rz -170.38 deg; joints [-12.476, 72.403, -175.69, 131.734, -60.838, 63.479, 2676.515, 474.819, 0]
  MoveL 189 to (743.95, -739.37, 869.23) mm, rotated rx 130.21 ry -8.72 rz -169.84 deg; joints [-12.476, 75.224, -179.751, 131.973, -60.065, 62.154, 2654.218, 488.345, 0]
  MoveL 190 to (709.42, -732.04, 889.63) mm, rotated rx 133.19 ry -9.83 rz -169.7 deg; joints [-12.476, 79.053, -185.502, 133.645, -58.375, 59.225, 2632.238, 514.975, 0]
  MoveL 191 to (673.05, -724.2, 910.56) mm, rotated rx 134.82 ry -10.39 rz -169.71 deg; joints [-12.476, 81.857, -189.951, 134.999, -57.948, 57.058, 2605.927, 534.847, 0]
  MoveL 192 to (634.86, -716.35, 931.75) mm, rotated rx 135.84 ry -10.15 rz -170.29 deg; joints [-12.476, 84.07, -193.661, 136.805, -58.584, 54.965, 2569.677, 551.383, 0]
  MoveL 193 to (590.38, -706.67, 956.08) mm, rotated rx 134.93 ry -9.14 rz -170.95 deg; joints [-13.013, 85.36, -195.933, 138.055, -60.928, 54.432, 2520.708, 551.818, 0]
  MoveL 194 to (534.66, -694.63, 985.12) mm, rotated rx 133.18 ry -7.68 rz -171.9 deg; joints [-13.013, 86.447, -197.926, 138.708, -64.085, 54.194, 2454.494, 554.996, 0.002]
  MoveL 195 to (471.61, -681.29, 1016.78) mm, rotated rx 130.54 ry -5.99 rz -173.05 deg; joints [-13.013, 87.161, -199.282, 138.966, -67.883, 54.662, 2377.062, 555.261, 0.001]
  MoveL 196 to (405.16, -667.16, 1047.91) mm, rotated rx 124.82 ry -2.46 rz -176.48 deg; joints [-12.982, 84.421, -199.282, 140.33, -77.278, 54.915, 2286.095, 552.193, 2.626]
  MoveL 197 to (341.85, -654.08, 1076.43) mm, rotated rx 122.99 ry -1.83 rz -177.19 deg; joints [-12.982, 85.194, -200.802, 140.238, -79.759, 55.286, 2218.458, 559.632, 0.082]
  MoveL 198 to (288.22, -643.1, 1099.97) mm, rotated rx 124.74 ry -1.97 rz -177.17 deg; joints [-12.982, 87.676, -206.184, 141.414, -80.688, 52.498, 2181.903, 582.709, 0]
  MoveL 199 to (239.56, -634.46, 1118.81) mm, rotated rx 128.95 ry 13.04 rz -164.09 deg; joints [-31.64, 82.162, -208.59, 150.889, -96.953, 37.959, 2259.037, 439.327, 0]
  MoveL 200 to (190.9, -627.66, 1133.72) mm, rotated rx 126.76 ry 14.31 rz -165.51 deg; joints [-31.64, 82.162, -208.589, 150.719, -99.462, 38.725, 2200.517, 438.925, 6.01]
  MoveL 201 to (142.76, -622.17, 1145.75) mm, rotated rx 124.74 ry 15.48 rz -167.01 deg; joints [-31.64, 82.162, -208.589, 150.763, -101.829, 39.458, 2141.901, 439.363, 13.545]
  MoveL 202 to (95.15, -617.72, 1156.22) mm, rotated rx 136.3 ry 27.91 rz -149.96 deg; joints [-44.422, 91.876, -166.166, 151.842, -57.295, 47.859, 1940.01, 93.218, 0.016]
  MoveL 203 to (45.18, -613.53, 1165.11) mm, rotated rx 140.79 ry 25.55 rz -147.99 deg; joints [-44.422, 95.911, -166.166, 150.356, -49.393, 48.719, 1870.377, 97.394, 0.001]
  MoveL 204 to (-9.5, -609.09, 1172.7) mm, rotated rx 137.9 ry 28.6 rz -150.73 deg; joints [-44.443, 95.606, -166.166, 152.95, -53.361, 47.699, 1800.439, 91.784, 22.931]
  MoveL 205 to (-66.79, -605.42, 1178.72) mm, rotated rx 136.64 ry 29.48 rz -151.63 deg; joints [-44.443, 95.632, -166.201, 153.428, -54.7, 47.81, 1739.995, 91.323, 29.345]
  MoveL 206 to (-124.09, -602.02, 1183.43) mm, rotated rx 133.51 ry 31.81 rz -154.34 deg; joints [-44.443, 95.508, -166.201, 155.176, -58.15, 47.675, 1671.169, 87.512, 54.709]
  MoveL 207 to (-178.76, -599.41, 1187.09) mm, rotated rx 133.6 ry 31.93 rz -154.49 deg; joints [-44.443, 95.508, -166.201, 155.436, -58.161, 47.456, 1614.474, 90.776, 51.361]
  MoveL 208 to (-228.21, -597.31, 1189.97) mm, rotated rx 133.46 ry 31.71 rz -154.21 deg; joints [-44.589, 95.508, -166.201, 155.135, -58.103, 47.789, 1570.121, 90.265, 47.767]
  MoveL 209 to (-273.47, -595.74, 1192.06) mm, rotated rx 136.82 ry 29.2 rz -151.33 deg; joints [-44.658, 95.507, -166.2, 153.394, -54.499, 47.837, 1538.388, 99.677, 11.784]
  MoveL 210 to (-315.85, -594.17, 1193.89) mm, rotated rx 141.11 ry 27.24 rz -149.49 deg; joints [-44.658, 97.542, -166.2, 152.858, -48.762, 47.23, 1485.019, 109.494, 0]
  MoveL 211 to (-357.71, -592.87, 1194.94) mm, rotated rx 138.48 ry 28.97 rz -151.11 deg; joints [-44.658, 97.414, -166.2, 153.623, -51.59, 47.611, 1439.228, 101.193, 21.649]
  MoveL 212 to (-400.87, -591.56, 1195.72) mm, rotated rx 133.78 ry 32.23 rz -154.85 deg; joints [-44.658, 96.97, -166.2, 155.938, -56.848, 47.556, 1383.279, 91.662, 61.038]
  MoveL 213 to (-447.44, -590.25, 1195.98) mm, rotated rx 135.87 ry 31.57 rz -153.98 deg; joints [-44.658, 96.707, -165.848, 156.176, -55.081, 46.59, 1333.576, 98.813, 43.206]
  MoveL 214 to (-498.72, -589.2, 1195.72) mm, rotated rx 138.74 ry 30.18 rz -152.35 deg; joints [-44.658, 96.655, -165.778, 155.89, -52.463, 45.673, 1283.852, 108.8, 19.418]
  MoveL 215 to (-560.72, -587.9, 1194.15) mm, rotated rx 138.79 ry 30.27 rz -152.44 deg; joints [-44.658, 96.577, -165.777, 156.086, -52.555, 45.483, 1220.948, 110.795, 20.377]
  MoveL 216 to (-639.47, -586.59, 1191.27) mm, rotated rx 142.52 ry 28.36 rz -150.48 deg; joints [-44.658, 97.182, -165.778, 155.693, -48.537, 44.439, 1141.12, 123.686, 0.003]
  MoveL 217 to (-727.63, -585.28, 1187.35) mm, rotated rx 144.41 ry 28.4 rz -150.44 deg; joints [-44.658, 97.542, -165.778, 157.123, -47.116, 42.604, 1041.244, 132.367, 0]
  MoveL 218 to (-817.62, -583.97, 1182.38) mm, rotated rx 148.91 ry 26.35 rz -148.6 deg; joints [-44.658, 99.834, -165.778, 156.95, -41.027, 41.319, 939.186, 145.924, 0]
  MoveL 219 to (-903.96, -583.19, 1176.36) mm, rotated rx 152.23 ry 24.86 rz -147.42 deg; joints [-44.738, 101.191, -165.778, 157.354, -36.865, 39.797, 845.179, 158.585, 0]
  MoveL 220 to (-980.87, -582.4, 1170.35) mm, rotated rx 154.34 ry 24.33 rz -146.96 deg; joints [-44.991, 101.599, -165.778, 158.922, -34.925, 37.667, 763.465, 166.916, 0]
  MoveL 221 to (-1045.23, -582.4, 1163.81) mm, rotated rx 157.67 ry 23.31 rz -146.16 deg; joints [-45.554, 102.479, -165.778, 161.669, -31.573, 34.101, 693.904, 177.207, 0]
  MoveL 222 to (-1093.1, -582.92, 1158.31) mm, rotated rx 160.05 ry 23.09 rz -145.83 deg; joints [-46.103, 102.703, -165.778, 165.192, -30.035, 30.105, 641.266, 183.81, 0]
  MoveL 223 to (-1127.38, -584.23, 1152.56) mm, rotated rx 159.19 ry 26.94 rz -147.87 deg; joints [-46.079, 100.059, -165.778, 170.003, -36.283, 26.091, 589.59, 183.81, 2.206]
  MoveL 224 to (-1150.66, -587.37, 1144.71) mm, rotated rx 155.94 ry 32.75 rz -152.02 deg; joints [-44.701, 99.059, -165.778, 172.164, -43.641, 25.274, 521.216, 184.543, 49.963]
  MoveL 225 to (-1167.93, -592.34, 1135.03) mm, rotated rx 153.43 ry 35.4 rz -154.59 deg; joints [-44.467, 96.744, -165.778, 173.427, -49.156, 25.326, 497.205, 184.543, 59.438]
  MoveL 226 to (-1183.88, -598.62, 1122.99) mm, rotated rx 151.57 ry 36.93 rz -156.37 deg; joints [-44.467, 94.397, -165.778, 174.26, -53.492, 25.506, 484.107, 184.541, 61.401]
  MoveL 227 to (-1198.01, -605.42, 1109.65) mm, rotated rx 148.78 ry 38.82 rz -158.96 deg; joints [-44.467, 91.959, -165.778, 175.138, -58.582, 26.153, 472.468, 184.54, 70.526]
  MoveL 228 to (-1209.26, -611.7, 1097.36) mm, rotated rx 147 ry 39.68 rz -160.44 deg; joints [-44.467, 90.097, -165.778, 175.416, -61.854, 26.747, 467.28, 184.54, 74.718]
  MoveL 229 to (-1219.72, -617.98, 1084.54) mm, rotated rx 144.88 ry 40.67 rz -162.27 deg; joints [-44.467, 88.389, -165.778, 175.791, -65.216, 27.456, 461.504, 184.539, 83.939]
  MoveL 230 to (-1231.24, -625.31, 1069.36) mm, rotated rx 143.52 ry 41.13 rz -163.31 deg; joints [-44.467, 86.674, -165.778, 175.885, -67.847, 27.962, 458.129, 184.539, 89.097]
  MoveL 231 to (-1243.79, -633.42, 1051.83) mm, rotated rx 141.86 ry 41.19 rz -164.05 deg; joints [-44.792, 85.593, -165.778, 175.682, -69.649, 28.964, 458.127, 174.356, 102.09]
  MoveL 232 to (-1258.18, -643.1, 1031.17) mm, rotated rx 140.7 ry 41.25 rz -164.59 deg; joints [-45.169, 84.091, -165.778, 175.755, -71.675, 29.544, 458.127, 166.68, 112.151]
  MoveL 233 to (-1272.83, -653.3, 1008.67) mm, rotated rx 138.47 ry 42.09 rz -166.6 deg; joints [-45.169, 82.243, -165.778, 176.203, -75.155, 30.26, 450.031, 166.68, 131.186]
  MoveL 234 to (-1285.91, -663.76, 985.65) mm, rotated rx 135.1 ry 43.09 rz -169.56 deg; joints [-45.169, 80.415, -165.778, 176.756, -79.265, 31.488, 442.666, 166.68, 157.811]
  MoveL 235 to (-1296.12, -673.97, 963.41) mm, rotated rx 132.2 ry 43.79 rz -172.12 deg; joints [-45.169, 78.832, -165.778, 177.232, -82.712, 32.573, 438.161, 166.68, 182.703]
  MoveL 236 to (-1301.61, -683.38, 943) mm, rotated rx 127.99 ry 44.17 rz -175.11 deg; joints [-45.438, 78.266, -165.778, 177.474, -85.57, 34.55, 438.159, 155.427, 220.19]
  MoveL 237 to (-1303.18, -692.02, 924.17) mm, rotated rx 122.92 ry 44.25 rz -178.39 deg; joints [-45.438, 79.694, -167.696, 177.195, -88.679, 37.059, 439.218, 142.971, 279.233]
  MoveL 238 to (-1301.87, -700.13, 907.16) mm, rotated rx 119.59 ry 44.04 rz 179.85 deg; joints [-45.679, 80.765, -169.148, 176.921, -90.687, 38.814, 447.599, 129.185, 323.312]
  MoveL 239 to (-1298.21, -707.71, 891.2) mm, rotated rx 116.95 ry 43.84 rz 178.45 deg; joints [-45.793, 81.677, -170.393, 176.678, -92.348, 40.182, 456.242, 118.579, 361.788]
  MoveL 240 to (-1292.98, -715.3, 876.03) mm, rotated rx 115.79 ry 43.72 rz 177.91 deg; joints [-45.906, 82.066, -170.927, 176.571, -93.064, 40.796, 464.8, 108.892, 386.659]
  MoveL 241 to (-1286.7, -722.36, 861.9) mm, rotated rx 114.7 ry 43.24 rz 178.49 deg; joints [-47.024, 82.267, -171.179, 176.426, -93.438, 41.67, 490.95, 85.22, 406.365]
  MoveL 242 to (-1279.63, -729.69, 848.04) mm, rotated rx 114.07 ry 43.06 rz 178.56 deg; joints [-47.421, 82.432, -171.406, 176.355, -93.755, 42.093, 505.529, 72.113, 424.568]
  MoveL 243 to (-1272.05, -736.49, 834.7) mm, rotated rx 114.85 ry 43.1 rz 179 deg; joints [-47.361, 82.006, -171.406, 176.355, -93.755, 41.68, 514.409, 69.006, 429.679]
  Set speed (1000.0 mm/s)
  MoveL 244 to (-1272.05, -736.49, 834.7) mm, rotated rx 114.85 ry 43.1 rz 179 deg; joints [-47.361, 82.006, -171.406, 176.355, -93.755, 41.68, 514.409, 69.006, 429.679]
  MoveL 245 to (-1302.34, -826.72, 865.38) mm, rotated rx 114.85 ry 43.1 rz 179 deg; joints [-47.361, 82.006, -171.406, 176.355, -93.755, 41.68, 484.114, -21.221, 398.996]

--- program Main_Prog (robot ABB IRB 1300-10/1.15) ---
  Set speed (1000.0 mm/s)
  MoveJ (Home)
  Call BumperR_C
  MoveJ (BumperR_Retreat)
  MoveJ (Trunk_App)
  Call Trunk_C
  Call Trunk_Top_C
  Call Top2_C
  MoveJ (Top_Retreat)
  MoveJ (Bonnet_App)
  Call Bonnet
  Call BumperF_C
  Call DoorFL_C
  Call DoorRL_C
  Call FrameL_C
  MoveJ (FrameL_Retreat)
  MoveJ (Front_Move)
  Call DoorFR_C
  Call DoorRR_C
  MoveJ (DoorRR_Retreat)
  Call FrameR_C
  MoveJ (Home)

--- program DoorRR (robot ABB IRB 1300-10/1.15) ---
  Smooth(1)
  Set speed (1000.0 mm/s)
  Set Ref.: DoorRR
  Set Tool: Generic Paint Sprayer
  Show Generic Paint Sprayer
  MoveJ 1 to (-63.47, 907.08, 255.99) mm, rotated rx 39.6 ry -2.99 rz 87.24 deg; joints [-128.12, 34.671, -33.35, 123.573, 79.803, -211.755, 1679.755, -179.592, 100.569]
  MoveL 2 to (-63.47, 907.08, 255.99) mm, rotated rx 39.6 ry -2.99 rz 87.24 deg; joints [-128.12, 34.671, -33.35, 123.573, 79.803, -211.755, 1679.757, -179.593, 100.574]
  MoveL 3 to (0, 900, 332.94) mm, rotated rx 39.6 ry -2.99 rz 87.24 deg; joints [-127.915, 34.535, -33.35, 123.577, 79.558, -211.755, 1679.759, -103.507, 162.351]
  MoveL 4 to (0, 900, 332.94) mm, rotated rx 39.6 ry -2.99 rz 87.24 deg; joints [-127.915, 34.535, -33.35, 123.577, 79.558, -211.755, 1679.759, -103.507, 162.351]
  Set speed (200.0 mm/s)
  MoveL 5 to (0, 800, 323.94) mm, rotated rx 38.28 ry -2.84 rz 87.41 deg; joints [-127.915, 34.519, -33.35, 122.717, 78.783, -210.888, 1781.675, -117.398, 172.973]
  MoveL 6 to (0, 700, 315.56) mm, rotated rx 37.73 ry -2.69 rz 87.55 deg; joints [-127.915, 34.519, -33.35, 122.423, 78.367, -210.547, 1883.605, -126.592, 178.774]
  MoveL 7 to (0, 600, 307.63) mm, rotated rx 36.98 ry -2.66 rz 87.59 deg; joints [-127.915, 34.516, -33.35, 121.882, 78.004, -210.043, 1984.114, -135.826, 186.427]
  MoveL 8 to (0, 500, 300.04) mm, rotated rx 32.16 ry -2.81 rz 87.64 deg; joints [-127.915, 34.515, -33.133, 118.177, 76.235, -206.887, 2083.534, -163.643, 224.679]
  MoveL 9 to (0, 400, 292.72) mm, rotated rx 31.37 ry -2.7 rz 87.73 deg; joints [-127.915, 34.515, -33.133, 117.621, 75.809, -206.341, 2184.841, -172.291, 232.801]
  MoveL 10 to (0, 300, 285.76) mm, rotated rx 30.76 ry -2.51 rz 87.86 deg; joints [-127.915, 34.515, -33.133, 117.245, 75.373, -205.932, 2286.918, -180.036, 239.468]
  MoveL 11 to (0, 200, 279.5) mm, rotated rx 29.26 ry -2.34 rz 87.99 deg; joints [-127.915, 34.515, -33.133, 116.14, 74.636, -204.876, 2388.784, -190.713, 252.814]
  MoveL 12 to (0, 100, 273.72) mm, rotated rx 28.63 ry -2.21 rz 88.07 deg; joints [-127.915, 34.515, -33.133, 115.701, 74.269, -204.437, 2490.209, -196.947, 259.916]
  MoveL 13 to (0, 0, 268.4) mm, rotated rx 25.03 ry -2.21 rz 88.12 deg; joints [-127.915, 34.514, -33.133, 112.751, 73.035, -201.769, 2590.477, -213.484, 290.009]
  Set speed (1000.0 mm/s)
  MoveL 14 to (0, 0, 268.4) mm, rotated rx 25.03 ry -2.21 rz 88.12 deg; joints [-127.915, 34.514, -33.133, 112.751, 73.035, -201.769, 2590.477, -213.484, 290.009]
  MoveL 15 to (-42.18, 4.87, 177.86) mm, rotated rx 25.03 ry -2.21 rz 88.12 deg; joints [-128.003, 34.551, -33.133, 112.748, 73.13, -201.769, 2590.477, -303.537, 248.292]
  Set speed (1000.0 mm/s)
  MoveL 16 to (77.33, 5.4, 118.5) mm, rotated rx -1.25 ry -3.13 rz 88.47 deg; joints [-131.414, 29.408, -33.133, 87.7, 73.13, -175.081, 2590.477, -334.567, 520.202]
  MoveL 17 to (75, 0, 218.33) mm, rotated rx -1.25 ry -3.13 rz 88.47 deg; joints [-131.159, 29.418, -33.133, 87.684, 72.876, -175.081, 2590.478, -237.209, 518.043]
  MoveL 18 to (75, 0, 218.33) mm, rotated rx -1.25 ry -3.13 rz 88.47 deg; joints [-131.159, 29.418, -33.133, 87.684, 72.876, -175.081, 2590.478, -237.209, 518.043]
  Set speed (200.0 mm/s)
  MoveL 19 to (75, 100, 223.81) mm, rotated rx 2.71 ry -3.1 rz 88.36 deg; joints [-131.372, 30.115, -33.133, 91.43, 72.876, -178.92, 2497.581, -237.209, 490.363]
  MoveL 20 to (75, 200, 229.45) mm, rotated rx 2.7 ry -3.22 rz 88.36 deg; joints [-131.372, 30.326, -33.133, 91.488, 73.005, -179.133, 2397.813, -235.278, 490.363]
  MoveL 21 to (75, 300, 235.32) mm, rotated rx 8.08 ry -3.19 rz 88.2 deg; joints [-131.372, 31.343, -33.133, 96.576, 73.203, -184.409, 2304.322, -235.278, 454.993]
  MoveL 22 to (75, 400, 241.4) mm, rotated rx 8.19 ry -3.31 rz 88.18 deg; joints [-131.372, 31.625, -33.133, 96.747, 73.362, -184.784, 2204.989, -233.26, 454.993]
  MoveL 23 to (75, 500, 247.79) mm, rotated rx 9.22 ry -3.43 rz 88.13 deg; joints [-131.372, 32.415, -33.133, 97.876, 73.675, -186.401, 2108.691, -233.26, 453.753]
  MoveL 24 to (75, 600, 261.44) mm, rotated rx 23.66 ry -23.77 rz 79.03 deg; joints [-131.372, 36.733, -33.133, 102.062, 97.93, -199.637, 1868.867, -104.915, 453.752]
  MoveL 25 to (75, 700, 280.68) mm, rotated rx 20.02 ry -2.78 rz 87.99 deg; joints [-140.774, 36.733, -29.31, 107.647, 86.181, -199.637, 2042.676, -104.915, 444.348]
  MoveL 26 to (75, 800, 276.44) mm, rotated rx 22.59 ry 10.54 rz 93.42 deg; joints [-143.982, 36.733, -29.31, 113.947, 76.326, -200.447, 2102.82, -104.915, 407.634]
  MoveL 27 to (75, 900, 278.65) mm, rotated rx -15.68 ry -40.48 rz 98.44 deg; joints [-134.388, 36.733, -29.31, 82.197, 113.909, -178.747, 1521.455, 43.242, 652.984]
  Set speed (1000.0 mm/s)
  MoveL 28 to (75, 900, 278.65) mm, rotated rx -15.68 ry -40.48 rz 98.44 deg; joints [-134.388, 36.733, -29.31, 82.197, 113.909, -178.747, 1521.455, 43.242, 652.984]
  MoveL 29 to (92.55, 965.79, 205.41) mm, rotated rx -15.68 ry -40.48 rz 98.44 deg; joints [-140.37, 35.88, -29.31, 81.467, 119.907, -178.747, 1517.07, 43.241, 657.394]
  Set speed (1000.0 mm/s)
  MoveL 30 to (120.12, 805.44, 147.11) mm, rotated rx 17.49 ry -2.67 rz 88.08 deg; joints [-161.484, 35.88, -29.31, 103.644, 105.044, -192.17, 2094.235, 43.241, 495.486]
  MoveL 31 to (150, 800, 242.38) mm, rotated rx 17.49 ry -2.67 rz 88.08 deg; joints [-161.185, 35.808, -29.31, 103.678, 104.739, -192.17, 2094.235, 134.311, 524.444]
  MoveL 32 to (150, 800, 242.38) mm, rotated rx 17.49 ry -2.67 rz 88.08 deg; joints [-161.185, 35.808, -29.31, 103.678, 104.739, -192.17, 2094.235, 134.311, 524.444]
  Set speed (200.0 mm/s)
  MoveL 33 to (150, 700, 237.54) mm, rotated rx 14.66 ry -1.9 rz 88.34 deg; joints [-161.654, 33.92, -29.31, 101.832, 103.527, -189.285, 2188.918, 134.311, 524.444]
  MoveL 34 to (150, 600, 232.62) mm, rotated rx 12 ry -2.62 rz 88.21 deg; joints [-161.609, 31.991, -29.31, 99.847, 103.527, -186.551, 2266.679, 134.311, 525.169]
  MoveL 35 to (150, 500, 227.36) mm, rotated rx 11.17 ry -2.76 rz 88.2 deg; joints [-161.667, 31.223, -29.31, 99.289, 103.527, -185.506, 2359.264, 133.93, 525.169]
  MoveL 36 to (150, 400, 221.99) mm, rotated rx 13.97 ry -2.53 rz 88.19 deg; joints [-161.642, 31.223, -29.31, 101.759, 103.527, -186.378, 2461.132, 135.141, 504.462]
  MoveL 37 to (150, 300, 216.85) mm, rotated rx 13.48 ry -2.49 rz 88.21 deg; joints [-161.788, 30.69, -29.31, 101.465, 103.47, -185.658, 2557.701, 135.141, 504.462]
  MoveL 38 to (150, 200, 211.93) mm, rotated rx 12.77 ry -2.29 rz 88.27 deg; joints [-161.959, 30.018, -29.31, 101.027, 103.254, -184.725, 2654.374, 135.141, 504.462]
  MoveL 39 to (150, 100, 207.2) mm, rotated rx 12.8 ry -2.35 rz 88.25 deg; joints [-161.959, 29.816, -29.31, 101.098, 103.27, -184.532, 2752.185, 133.949, 504.462]
  MoveL 40 to (150, 0, 203.02) mm, rotated rx 12.74 ry -1.88 rz 88.36 deg; joints [-162.195, 29.772, -29.31, 101.098, 103.011, -184.412, 2857.032, 133.949, 506.753]
  Set speed (1000.0 mm/s)
  MoveL 41 to (150, 0, 203.02) mm, rotated rx 12.74 ry -1.88 rz 88.36 deg; joints [-162.195, 29.772, -29.31, 101.098, 103.011, -184.412, 2857.032, 133.949, 506.753]
  MoveL 42 to (128.05, 3.83, 105.54) mm, rotated rx 12.74 ry -1.88 rz 88.36 deg; joints [-162.291, 29.791, -29.31, 101.097, 103.109, -184.412, 2857.031, 37.709, 485.046]
  Set speed (1000.0 mm/s)
  MoveL 43 to (220.65, 4.01, 93.86) mm, rotated rx 2.55 ry -2.23 rz 88.41 deg; joints [-162.381, 29.791, -29.31, 92.09, 103.109, -181.268, 2852.075, 17.236, 664.089]
  MoveL 44 to (225, 0, 193.68) mm, rotated rx 2.55 ry -2.23 rz 88.41 deg; joints [-162.381, 29.79, -29.31, 92.09, 103.109, -181.268, 2853.288, 117.133, 668.44]
  MoveL 45 to (225, 0, 193.68) mm, rotated rx 2.55 ry -2.23 rz 88.41 deg; joints [-162.381, 29.79, -29.31, 92.09, 103.109, -181.268, 2853.288, 117.133, 668.44]
  Set speed (200.0 mm/s)
  MoveL 46 to (225, 100, 197.78) mm, rotated rx 2.48 ry -2.34 rz 88.4 deg; joints [-162.275, 29.891, -29.31, 92.001, 103.109, -181.353, 2752.783, 117.133, 667.602]
  MoveL 47 to (225, 200, 202.17) mm, rotated rx 2.48 ry -2.51 rz 88.4 deg; joints [-162.105, 29.891, -29.31, 91.999, 103.117, -181.361, 2650.435, 117.134, 664.884]
  MoveL 48 to (225, 300, 206.77) mm, rotated rx 2.74 ry -2.52 rz 88.39 deg; joints [-162.081, 30.282, -29.31, 92.128, 103.117, -181.841, 2553.676, 117.697, 664.884]
  MoveL 49 to (225, 400, 211.28) mm, rotated rx 3.42 ry -2.45 rz 88.38 deg; joints [-162.087, 30.966, -29.31, 92.575, 103.105, -182.758, 2460.23, 117.697, 664.884]
  MoveL 50 to (225, 500, 215.72) mm, rotated rx 3.72 ry -2.47 rz 88.38 deg; joints [-162.033, 31.38, -29.31, 92.737, 103.105, -183.277, 2363.307, 117.767, 664.884]
  MoveL 51 to (225, 600, 220.75) mm, rotated rx 5.54 ry -1.67 rz 88.42 deg; joints [-162.275, 32.835, -29.31, 94.068, 102.758, -185.308, 2283.425, 117.768, 664.883]
  MoveL 52 to (225, 700, 223.76) mm, rotated rx 6.11 ry -1.55 rz 88.44 deg; joints [-162.343, 33.331, -29.31, 94.465, 102.783, -185.981, 2188.915, 117.767, 663.691]
  Set speed (1000.0 mm/s)
  MoveL 53 to (225, 700, 223.76) mm, rotated rx 6.11 ry -1.55 rz 88.44 deg; joints [-162.343, 33.331, -29.31, 94.465, 102.783, -185.981, 2188.915, 117.767, 663.691]
  MoveL 54 to (214.44, 702.97, 124.36) mm, rotated rx 6.11 ry -1.55 rz 88.44 deg; joints [-162.344, 33.331, -29.31, 94.464, 102.784, -185.981, 2188.908, 18.351, 653.156]
  Set speed (1000.0 mm/s)
  MoveL 55 to (297.16, 702.27, 119.51) mm, rotated rx 1.66 ry -1.26 rz 88.45 deg; joints [-162.845, 32.919, -29.31, 90.621, 102.636, -184.182, 2188.908, 18.351, 768.606]
  MoveL 56 to (300, 700, 219.45) mm, rotated rx 1.66 ry -1.26 rz 88.45 deg; joints [-162.845, 32.919, -29.31, 90.621, 102.636, -184.182, 2188.421, 118.31, 771.407]
  MoveL 57 to (300, 700, 219.45) mm, rotated rx 1.66 ry -1.26 rz 88.45 deg; joints [-162.845, 32.919, -29.31, 90.621, 102.636, -184.182, 2188.421, 118.31, 771.407]
  Set speed (200.0 mm/s)
  MoveL 58 to (300, 600, 217.1) mm, rotated rx -0.28 ry -1.56 rz 88.44 deg; joints [-162.631, 31.395, -29.31, 89.23, 102.636, -182.032, 2271.976, 120.497, 771.408]
  MoveL 59 to (300, 500, 213.93) mm, rotated rx -0.88 ry -1.74 rz 88.44 deg; joints [-162.497, 30.775, -29.31, 88.842, 102.674, -181.213, 2364.505, 120.497, 771.408]
  MoveL 60 to (300, 400, 210.18) mm, rotated rx -0.47 ry -2.5 rz 88.45 deg; joints [-162.359, 30.775, -29.31, 89.186, 103.308, -181.34, 2457.368, 120.497, 770.637]
  MoveL 61 to (300, 300, 205.93) mm, rotated rx -1.36 ry -2.52 rz 88.46 deg; joints [-162.34, 29.951, -29.31, 88.599, 103.308, -180.217, 2549.963, 121.143, 770.638]
  MoveL 62 to (300, 200, 201.56) mm, rotated rx -1.07 ry -2.61 rz 88.46 deg; joints [-162.34, 29.932, -29.31, 88.859, 103.403, -180.287, 2649.035, 119.839, 770.638]
  MoveL 63 to (300, 100, 197.15) mm, rotated rx -0.69 ry -2.46 rz 88.45 deg; joints [-162.486, 29.932, -29.31, 89.194, 103.403, -180.408, 2751.005, 119.554, 770.123]
  MoveL 64 to (300, 0, 193.08) mm, rotated rx -2.06 ry -2.36 rz 88.47 deg; joints [-162.486, 28.762, -29.31, 88.262, 103.336, -178.782, 2841.368, 121.371, 770.126]
  Set speed (1000.0 mm/s)
  MoveL 65 to (300, 0, 193.08) mm, rotated rx -2.06 ry -2.36 rz 88.47 deg; joints [-162.486, 28.762, -29.31, 88.262, 103.336, -178.782, 2841.368, 121.371, 770.126]
  MoveL 66 to (303.7, 4.02, 93.23) mm, rotated rx -2.06 ry -2.36 rz 88.47 deg; joints [-162.486, 28.762, -29.31, 88.262, 103.336, -178.782, 2839.932, 21.451, 773.819]
  Set speed (1000.0 mm/s)
  MoveL 67 to (382.7, 3.94, 97.57) mm, rotated rx -4.36 ry -2.38 rz 88.5 deg; joints [-162.412, 28.762, -29.31, 86.236, 103.336, -178.068, 2837.249, 25.97, 872.373]
  MoveL 68 to (375, 0, 197.2) mm, rotated rx -4.36 ry -2.38 rz 88.5 deg; joints [-162.412, 28.762, -29.31, 86.236, 103.336, -178.068, 2838.719, 125.661, 864.677]
  MoveL 69 to (375, 0, 197.2) mm, rotated rx -4.36 ry -2.38 rz 88.5 deg; joints [-162.412, 28.762, -29.31, 86.236, 103.336, -178.068, 2838.719, 125.661, 864.677]
  Set speed (200.0 mm/s)
  MoveL 70 to (375, 100, 201.22) mm, rotated rx -4.3 ry -2.5 rz 88.51 deg; joints [-162.336, 29.015, -29.31, 86.228, 103.366, -178.339, 2739.592, 125.662, 864.558]
  MoveL 71 to (375, 200, 205.44) mm, rotated rx -4.44 ry -2.52 rz 88.51 deg; joints [-162.318, 29.145, -29.31, 86.081, 103.366, -178.429, 2640.442, 126.742, 864.557]
  MoveL 72 to (375, 300, 209.49) mm, rotated rx -3.68 ry -2.33 rz 88.49 deg; joints [-162.457, 29.879, -29.31, 86.564, 103.249, -179.426, 2549.304, 126.742, 864.556]
  MoveL 73 to (375, 400, 213.08) mm, rotated rx -3.23 ry -2.01 rz 88.46 deg; joints [-162.601, 30.402, -29.31, 86.837, 103.043, -180.109, 2457.26, 126.742, 864.556]
  MoveL 74 to (375, 500, 216.05) mm, rotated rx -2.67 ry -1.73 rz 88.45 deg; joints [-162.789, 30.998, -29.31, 87.195, 102.922, -180.903, 2365.744, 126.742, 864.556]
  MoveL 75 to (375, 600, 218.52) mm, rotated rx -1.86 ry -1.36 rz 88.43 deg; joints [-163.06, 31.755, -29.31, 87.734, 102.806, -181.932, 2276.656, 126.742, 864.555]
  Set speed (1000.0 mm/s)
  MoveL 76 to (375, 600, 218.52) mm, rotated rx -1.86 ry -1.36 rz 88.43 deg; joints [-163.06, 31.755, -29.31, 87.734, 102.806, -181.932, 2276.656, 126.742, 864.555]
  MoveL 77 to (378.31, 602.28, 118.6) mm, rotated rx -1.86 ry -1.36 rz 88.43 deg; joints [-163.06, 31.719, -29.31, 87.742, 102.807, -181.895, 2276.656, 26.893, 867.444]
  Set speed (1000.0 mm/s)
  MoveL 78 to (454.83, 601.84, 122) mm, rotated rx -2.74 ry -1.13 rz 88.42 deg; joints [-163.06, 31.69, -29.31, 86.972, 102.556, -181.6, 2276.657, 29.818, 951.2]
  MoveL 79 to (450, 600, 221.87) mm, rotated rx -2.74 ry -1.13 rz 88.42 deg; joints [-163.06, 31.773, -29.31, 86.954, 102.551, -181.685, 2276.656, 129.48, 947.372]
  MoveL 80 to (450, 600, 221.87) mm, rotated rx -2.74 ry -1.13 rz 88.42 deg; joints [-163.06, 31.773, -29.31, 86.954, 102.551, -181.685, 2276.656, 129.48, 947.372]
  Set speed (200.0 mm/s)
  MoveL 81 to (450, 500, 220.16) mm, rotated rx -3.81 ry -0.92 rz 88.4 deg; joints [-163.06, 30.826, -29.31, 86.215, 102.377, -180.396, 2370.308, 132.655, 947.373]
  MoveL 82 to (450, 400, 218.21) mm, rotated rx -4.34 ry -1.74 rz 88.45 deg; joints [-162.66, 30.264, -29.31, 85.883, 102.838, -179.631, 2456.489, 132.655, 947.374]
  MoveL 83 to (450, 300, 215.34) mm, rotated rx -4.61 ry -1.94 rz 88.47 deg; joints [-162.526, 29.864, -29.31, 85.74, 102.939, -179.129, 2550.615, 132.655, 947.374]
  MoveL 84 to (450, 200, 211.78) mm, rotated rx -4.24 ry -2.17 rz 88.48 deg; joints [-162.526, 29.864, -29.31, 86.077, 103.169, -179.244, 2648.628, 132.472, 946.812]
  MoveL 85 to (450, 100, 207.82) mm, rotated rx -4.65 ry -2.42 rz 88.51 deg; joints [-162.426, 29.366, -29.31, 85.837, 103.362, -178.599, 2741.604, 132.472, 946.812]
  MoveL 86 to (450, 0, 203.99) mm, rotated rx -4.99 ry -2.31 rz 88.5 deg; joints [-162.431, 28.907, -29.31, 85.643, 103.291, -178.024, 2838.512, 132.472, 946.812]
  Set speed (1000.0 mm/s)
  MoveL 87 to (450, 0, 203.99) mm, rotated rx -4.99 ry -2.31 rz 88.5 deg; joints [-162.431, 28.907, -29.31, 85.643, 103.291, -178.024, 2838.512, 132.472, 946.812]
  MoveL 88 to (458.8, 3.78, 104.45) mm, rotated rx -4.99 ry -2.31 rz 88.5 deg; joints [-162.431, 28.907, -29.31, 85.643, 103.291, -178.024, 2837.167, 32.868, 955.604]
  Set speed (1000.0 mm/s)
  MoveL 89 to (515.12, 3.49, 104.06) mm, rotated rx 5.73 ry -1.85 rz 88.41 deg; joints [-162.551, 28.907, -29.31, 95.108, 102.904, -181.329, 2840.382, 32.868, 920.358]
  MoveL 90 to (525, 0, 203.5) mm, rotated rx 5.73 ry -1.85 rz 88.41 deg; joints [-162.551, 28.907, -29.31, 95.108, 102.904, -181.329, 2840.929, 132.377, 930.229]
  MoveL 91 to (525, 0, 203.5) mm, rotated rx 5.73 ry -1.85 rz 88.41 deg; joints [-162.551, 28.907, -29.31, 95.108, 102.904, -181.329, 2840.929, 132.377, 930.229]
  Set speed (200.0 mm/s)
  MoveL 92 to (525, 100, 207.22) mm, rotated rx 5.48 ry -2.06 rz 88.39 deg; joints [-162.441, 28.953, -29.31, 94.874, 103.008, -181.312, 2738.998, 132.377, 930.229]
  MoveL 93 to (525, 200, 211.32) mm, rotated rx 5.33 ry -2.41 rz 88.36 deg; joints [-162.259, 28.983, -29.31, 94.718, 103.169, -181.312, 2635.468, 132.377, 929.32]
  MoveL 94 to (525, 300, 215.9) mm, rotated rx 5.32 ry -2.56 rz 88.34 deg; joints [-162.095, 29.055, -29.31, 94.686, 103.169, -181.397, 2533.967, 132.377, 927.595]
  MoveL 95 to (525, 400, 220.62) mm, rotated rx 3.08 ry -2.6 rz 88.38 deg; joints [-162.094, 29.055, -29.31, 92.712, 103.169, -180.69, 2433.601, 133.162, 943.953]
  MoveL 96 to (525, 500, 224.64) mm, rotated rx 0.01 ry -1.71 rz 88.44 deg; joints [-162.302, 29.055, -29.31, 90.017, 102.478, -179.724, 2342.137, 133.162, 967.298]
  Set speed (1000.0 mm/s)
  MoveL 97 to (525, 500, 224.64) mm, rotated rx 0.01 ry -1.71 rz 88.44 deg; joints [-162.302, 29.055, -29.31, 90.017, 102.478, -179.724, 2342.137, 133.162, 967.298]
  MoveL 98 to (525.06, 502.99, 124.68) mm, rotated rx 0.01 ry -1.71 rz 88.44 deg; joints [-162.302, 29.055, -29.31, 90.017, 102.478, -179.724, 2341.831, 33.165, 967.376]

